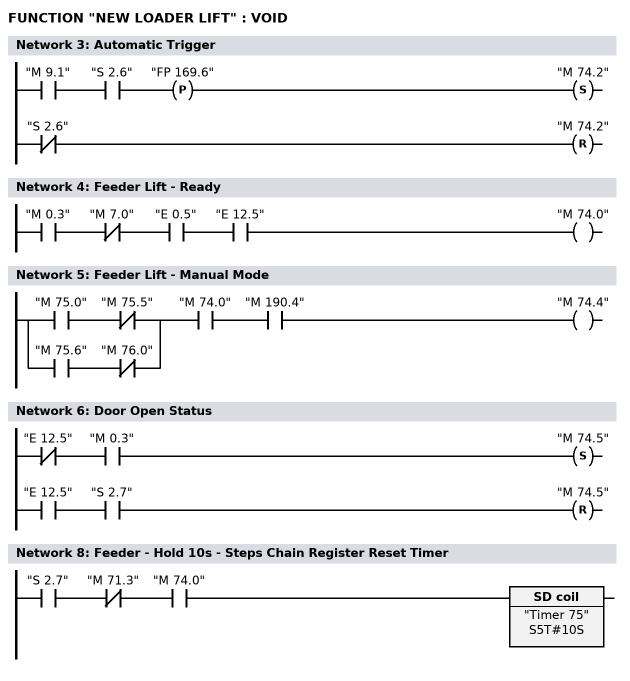

      O     "M 9.1";
      A     "S 2.6";
      FP    "FP 169.6";
      S     "M 74.2";
//;
      AN    "S 2.6";
      R     "M 74.2";
NETWORK
TITLE =Feeder Lift - Ready

      A     "M 0.3";
      AN    "M 7.0";
      A     "E 0.5";
      A     "E 12.5";
      =     "M 74.0";
NETWORK
TITLE =Feeder Lift - Manual Mode

      A(    ;
      A     "M 75.0";
      AN    "M 75.5";
      O     ;
      A     "M 75.6";
      AN    "M 76.0";
      )     ;
      A     "M 74.0";
      A     "M 190.4";
      =     "M 74.4";
NETWORK
TITLE =Door Open Status

      AN    "E 12.5";
      A     "M 0.3";
      S     "M 74.5";
//;
      A     "E 12.5";
      A     "S 2.7";
      R     "M 74.5";
NETWORK
TITLE =Fault Reset Status        X121     transfered to FC 212 Net 79
//      A(
//      O     "M 54.7"
//      O     "M 66.7"
//      O     "M 86.7"
//      )
//      A     "M 145.0"
//      O     "M 74.5"
//      O     "Timer 0"
//      =     "H 40.3"
//
//is transfered to FC 212 Net 79


NETWORK
TITLE =Feeder - Hold 10s - Steps Chain Register Reset Timer

      A     "S 2.7";
      AN    "M 71.3";
      A     "M 74.0";
      L     S5T#10S;
      SD    "Timer 75";
NETWORK
TITLE =Feeder - All Register Reset

      A(    ;
      A     "M 190.4";
      A     "M 171.4";
      A     "M 171.5";
      O     "Timer 75";
      )     ;
      A     "M 74.0";
      JC    M001;
      JU    M002;

M001: L     2#0;
      T     "MW 71";
      T     "MW 75";

M002: NOP   0;
NETWORK
TITLE =Step 16N1 - Power On
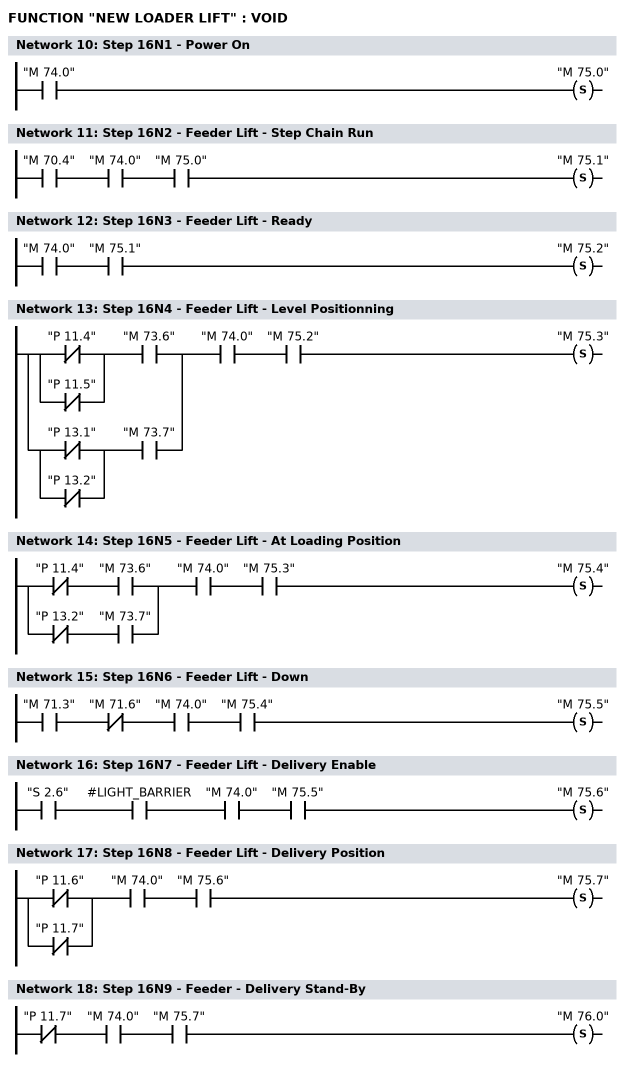

      A     "M 74.0";
      S     "M 75.0";
NETWORK
TITLE =Step 16N2 - Feeder Lift - Step Chain Run

      A     "M 70.4";
      A     "M 74.0";
      A     "M 75.0";
      S     "M 75.1";
NETWORK
TITLE =Step 16N3 - Feeder Lift - Ready

      A     "M 74.0";
      A     "M 75.1";
      S     "M 75.2";
NETWORK
TITLE =Step 16N4 - Feeder Lift - Level Positionning

      A(    ;
      A(    ;
      ON    "P 11.4";
      ON    "P 11.5";
      )     ;
      A     "M 73.6";
      O     ;
      A(    ;
      ON    "P 13.1";
      ON    "P 13.2";
      )     ;
      A     "M 73.7";
      )     ;
      A     "M 74.0";
      A     "M 75.2";
      S     "M 75.3";
NETWORK
TITLE =Step 16N5 - Feeder Lift - At Loading Position

      A(    ;
      AN    "P 11.4";
      A     "M 73.6";
      O     ;
      AN    "P 13.2";
      A     "M 73.7";
      )     ;
      A     "M 74.0";
      A     "M 75.3";
      S     "M 75.4";
NETWORK
TITLE =Step 16N6 - Feeder Lift - Down

      A     "M 71.3";
      AN    "M 71.6";
      A     "M 74.0";
      A     "M 75.4";
      S     "M 75.5";
NETWORK
TITLE =Step 16N7 - Feeder Lift - Delivery Enable

      A     "S 2.6";
      A     #LIGHT_BARRIER;
      A     "M 74.0";
      A     "M 75.5";
      S     "M 75.6";
NETWORK
TITLE =Step 16N8 - Feeder Lift - Delivery Position

      A(    ;
      ON    "P 11.6";
      ON    "P 11.7";
      )     ;
      A     "M 74.0";
      A     "M 75.6";
      S     "M 75.7";
NETWORK
TITLE =Step 16N9 - Feeder - Delivery Stand-By

      AN    "P 11.7";
      A     "M 74.0";
      A     "M 75.7";
      S     "M 76.0";
NETWORK
TITLE =Feeder Lift Steps Chain Reset by Feeder Fingers (MW71)

      A     "M 76.0";
      AN    "M 76.1";
      A(    ;
      ON    "M 71.2";
      O     "M 72.2";
      )     ;
      A     "M 74.0";
      JC    M003;
      JU    M004;

M003: L     2#0;
      T     "MW 75";

M004: NOP   0;
NETWORK
TITLE =Step 16N10 - Feeder Hold Operation (Stop) 1
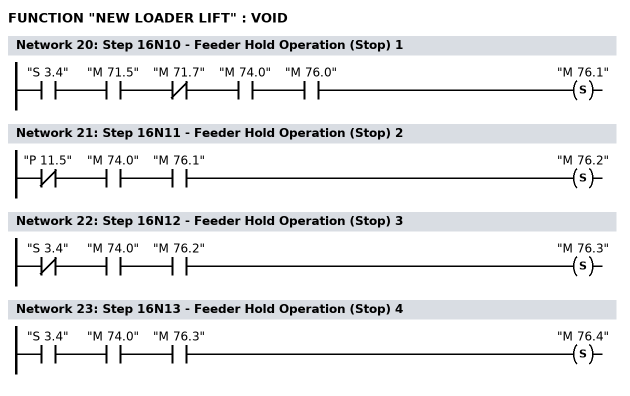

      A     "S 3.4";
      A     "M 71.5";
      AN    "M 71.7";
      A     "M 74.0";
      A     "M 76.0";
      S     "M 76.1";
NETWORK
TITLE =Step 16N11 - Feeder Hold Operation (Stop) 2

      AN    "P 11.5";
      A     "M 74.0";
      A     "M 76.1";
      S     "M 76.2";
NETWORK
TITLE =Step 16N12 - Feeder Hold Operation (Stop) 3

      AN    "S 3.4";
      A     "M 74.0";
      A     "M 76.2";
      S     "M 76.3";
NETWORK
TITLE =Step 16N13 - Feeder Hold Operation (Stop) 4

      A     "S 3.4";
      A     "M 74.0";
      A     "M 76.3";
      S     "M 76.4";
NETWORK
TITLE =Step 16N14 - Feeder Hold Operation (Stop) 4 - Fill MB76

      A     "M 76.4";
      A     "M 74.0";
      JC    M005;
      JU    M006;

M005: L     2#11111100000000;
      T     "MW 75";

M006: NOP   0;
NETWORK
TITLE =Packets Movements - UpDate
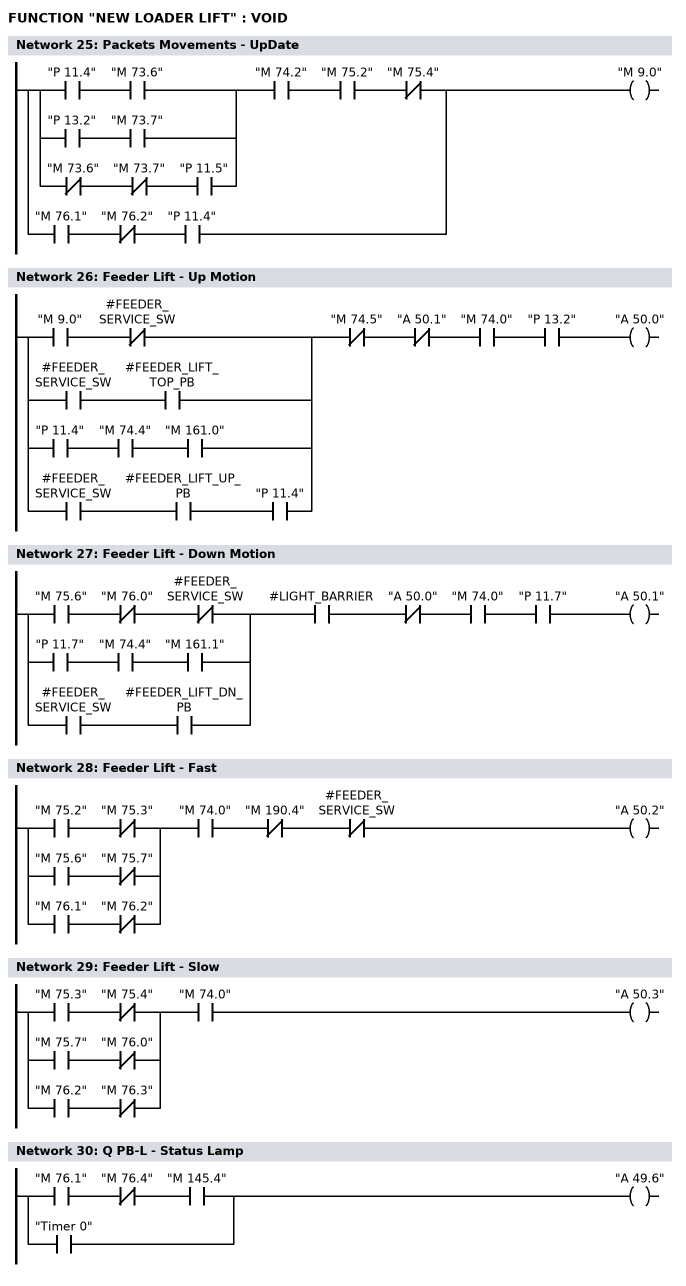

      A(    ;
      A     "P 11.4";
      A     "M 73.6";
      O     ;
      A     "P 13.2";
      A     "M 73.7";
      O     ;
      AN    "M 73.6";
      AN    "M 73.7";
      A     "P 11.5";
      )     ;
      A     "M 74.2";
      A     "M 75.2";
      AN    "M 75.4";
      O     ;
      A     "M 76.1";
      AN    "M 76.2";
      A     "P 11.4";
      =     "M 9.0";
NETWORK
TITLE =Feeder Lift - Up Motion

      A(    ;
      A     "M 9.0";
      AN    #FEEDER_SERVICE_SW;
      O     ;
      A     #FEEDER_SERVICE_SW;
      A     #FEEDER_LIFT_TOP_PB;

      O     ;
      A     "P 11.4";
      A     "M 74.4";
      A     "M 161.0";

      O     ;
      A     #FEEDER_SERVICE_SW;
      A     #FEEDER_LIFT_UP_PB;
      A     "P 11.4";
      )     ;
      AN    "M 74.5";
      AN    "A 50.1";
      A     "M 74.0";
      A     "P 13.2";
      =     "A 50.0";
NETWORK
TITLE =Feeder Lift - Down Motion

      A(    ;
      A     "M 75.6";
      AN    "M 76.0";
      AN    #FEEDER_SERVICE_SW;

      O     ;
      A     "P 11.7";
      A     "M 74.4";
      A     "M 161.1";

      O     ;
      A     #FEEDER_SERVICE_SW;
      A     #FEEDER_LIFT_DN_PB;
      )     ;
      A     #LIGHT_BARRIER;
      AN    "A 50.0";
      A     "M 74.0";
      A     "P 11.7";
      =     "A 50.1";
NETWORK
TITLE =Feeder Lift - Fast

      A(    ;
      A     "M 75.2";
      AN    "M 75.3";
      O     ;
      A     "M 75.6";
      AN    "M 75.7";
      O     ;
      A     "M 76.1";
      AN    "M 76.2";
      )     ;
      A     "M 74.0";
      AN    "M 190.4";
      AN    #FEEDER_SERVICE_SW;
      =     "A 50.2";
NETWORK
TITLE =Feeder Lift - Slow

      A(    ;
      A     "M 75.3";
      AN    "M 75.4";
      O     ;
      A     "M 75.7";
      AN    "M 76.0";
      O     ;
      A     "M 76.2";
      AN    "M 76.3";
      )     ;
      A     "M 74.0";
      =     "A 50.3";
NETWORK
TITLE =Q PB-L - Status Lamp

      A     "M 76.1";
      AN    "M 76.4";
      A     "M 145.4";
      O     "Timer 0";
      =     "A 49.6";
END_FUNCTION

FUNCTION "NEW C21 - LINK 1 HI" : VOID
TITLE =NEW FC978 (was FC1078) - Conveyor 21 - Link 1H Pos. 13 High Leve
//
//v0.1 2026-11-19: clearing trigger M9.3 only if pivot HIGH (P15.0).
NAME : POS_13_H
VERSION : 0.1


VAR_TEMP
  MAIN_SERVICE_2_SW : BOOL ;
  SERVICE_RUN : BOOL ;
  INITIALISATION : BOOL ;
  BARRIER_BLINKER : BOOL ;
END_VAR
BEGIN
NETWORK
TITLE =Conveyor 21 - Service

      A     "HMI_DB".ALL_SERVICE_ENABLE_SW;
      A     "HMI_DB".CONVEYOR_21_SERVICE_SW;
      A     "HMI_DB".SERVICE_SW_2_STATUS;
      =     #MAIN_SERVICE_2_SW;
//;
      A     #MAIN_SERVICE_2_SW;
      O     "M 78.7";
      JNB   CO21;
//;
      A     "HMI_DB".HMI_CONVEYOR_21_TEST_SSW;
      AN    "A 48.0";
      =     #SERVICE_RUN;
      S     "DB UTILITY".Conveyor_10_Disable;
      S     "DB UTILITY".Pivot_Disable;
//;
      A     "HMI_DB".SERVICE_INIT_PB;
      =     #INITIALISATION;
//;
      AN    #MAIN_SERVICE_2_SW;
      R     "HMI_DB".HMI_CONVEYOR_21_TEST_SSW;
      R     "DB UTILITY".Conveyor_10_Disable;
      R     "DB UTILITY".Pivot_Disable;

CO21: R     #SERVICE_RUN;
      R     #INITIALISATION; // Fix: temp not written when service is off
      FP    "FP 148.3";
      =     "M 78.7";
NETWORK
TITLE =Power Enable
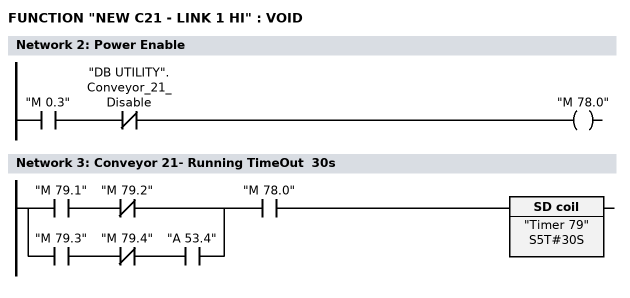

      A     "M 0.3";
      AN    "DB UTILITY".Conveyor_21_Disable;
      =     "M 78.0";
NETWORK
TITLE =Conveyor 21- Running TimeOut  30s

      A(    ;
      A     "M 79.1";
      AN    "M 79.2";
      O     ;
      A     "M 79.3";
      AN    "M 79.4";
      A     "A 53.4";
      )     ;
      A     "M 78.0";
      L     S5T#30S;
      SD    "Timer 79"; // C21 TimeOut
NETWORK
TITLE =Steps Register - Reset

      A(    ;
      A     "M 79.1"; // Filling Step
      AN    "M 79.2"; // Filling Step - Done
      A     "Timer 79"; // C21 TimeOut
      O     "M 79.4";
      O     #INITIALISATION;
      O     "DB UTILITY".Conveyor_21_Disable;
      )     ;
      A     "M 78.0";
      JC    M001;
      JU    M002;

M001: L     W#16#0;
      T     "MW 79"; // Step Register - Reset
      T     "MB 81"; // Step Register - Reset

M002: NOP   0;
NETWORK
TITLE =Step 22N1 - Power ON
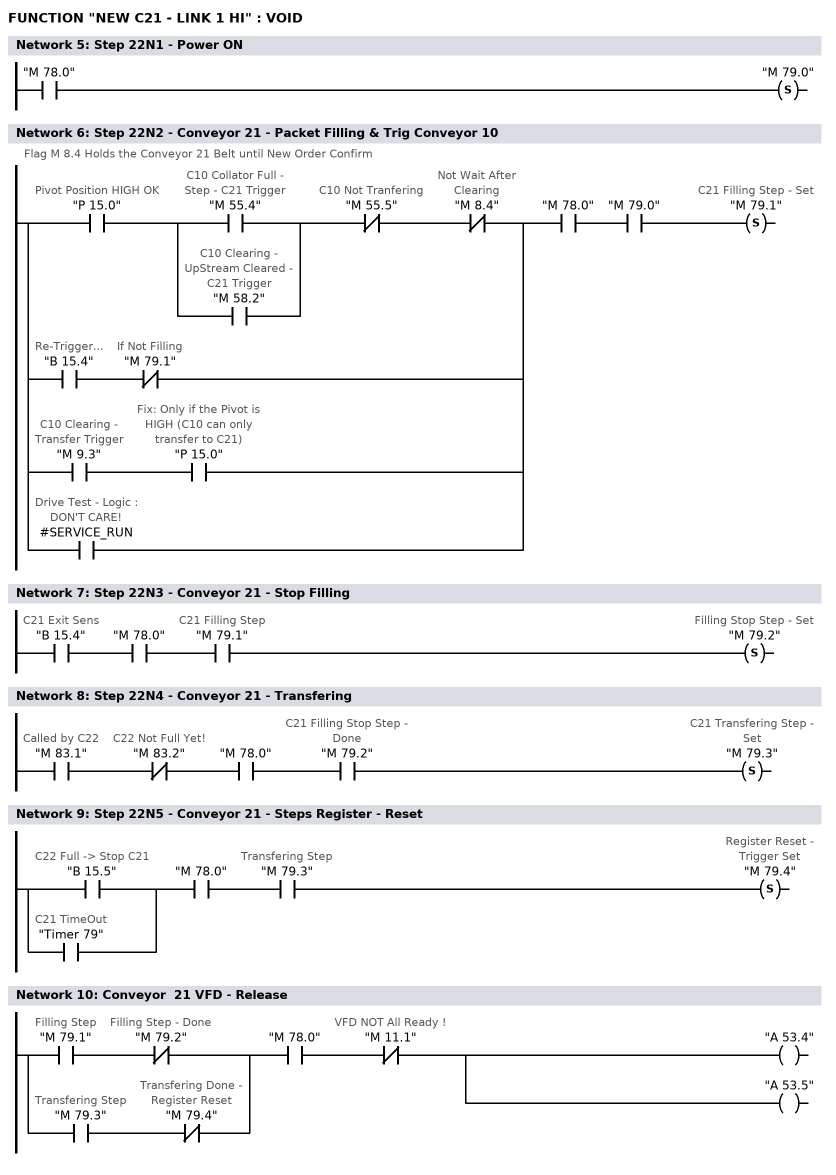

      A     "M 78.0";
      S     "M 79.0";
NETWORK
TITLE =Step 22N2 - Conveyor 21 - Packet Filling & Trig Conveyor 10
//Flag M 8.4 Holds the Conveyor 21 Belt until New Order Confirm
      A(    ;
      A     "P 15.0"; // Pivot Position HIGH OK
      A(    ;
      O     "M 55.4"; // C10 Collator Full - Step - C21 Trigger
      O     "M 58.2"; // C10 Clearing - UpStream Cleared - C21 Trigger
      )     ;
      AN    "M 55.5"; // C10 Not Tranfering
      AN    "M 8.4"; // Not Wait After Clearing
      O     ;
      A     "B 15.4"; // Re-Trigger...
      AN    "M 79.1"; // If Not Filling
      O     ;
      A     "M 9.3"; // C10 Clearing - Transfer Trigger
      A     "P 15.0"; // Fix: Only if the Pivot is HIGH (C10 can only transfer to C21)
      )     ;
      O     #SERVICE_RUN; // Drive Test - Logic : DON'T CARE!
      A     "M 78.0";
      A     "M 79.0";
      S     "M 79.1"; // C21 Filling Step - Set
NETWORK
TITLE =Step 22N3 - Conveyor 21 - Stop Filling

      A     "B 15.4"; // C21 Exit Sens
      A     "M 78.0";
      A     "M 79.1"; // C21 Filling Step
      S     "M 79.2"; // Filling Stop Step - Set
NETWORK
TITLE =Step 22N4 - Conveyor 21 - Transfering

      A     "M 83.1"; // Called by C22
      AN    "M 83.2"; // C22 Not Full Yet!
      A     "M 78.0";
      A     "M 79.2"; // C21 Filling Stop Step - Done
      S     "M 79.3"; // C21 Transfering Step - Set
NETWORK
TITLE =Step 22N5 - Conveyor 21 - Steps Register - Reset

      A(    ;
      O     "B 15.5"; // C22 Full -> Stop C21
      O     "Timer 79"; // C21 TimeOut
      )     ;
      A     "M 78.0";
      A     "M 79.3"; // Transfering Step
      S     "M 79.4"; // Register Reset - Trigger Set
NETWORK
TITLE =Conveyor  21 VFD - Release

      A(    ;
      A     "M 79.1"; // Filling Step
      AN    "M 79.2"; // Filling Step - Done
      O     ;
      A     "M 79.3"; // Transfering Step
      AN    "M 79.4"; // Transfering Done - Register Reset
      )     ;
      A     "M 78.0";
      AN    "M 11.1"; // VFD NOT All Ready !
      =     "A 53.4";
      =     "A 53.5";
END_FUNCTION

FUNCTION "NEW C22 - LINK 2 HI" : VOID
TITLE =NEW FC982 (was FC1082) - Conveyor 22 - Link 2H Pos. 14 High Leve
//
NAME : POS_14_H
VERSION : 0.0


VAR_TEMP
  MAIN_SERVICE_2_SW : BOOL ;
  SERVICE_RUN : BOOL ;
END_VAR
BEGIN
NETWORK
TITLE =Conveyor 22 - Service

      A     "HMI_DB".ALL_SERVICE_ENABLE_SW;
      A     "HMI_DB".CONVEYOR_21_SERVICE_SW;
      A     "HMI_DB".SERVICE_SW_2_STATUS;
      =     #MAIN_SERVICE_2_SW;
//;
      A     #MAIN_SERVICE_2_SW;
      O     "M 82.7";
      JNB   CO22;
//;
      A     "HMI_DB".HMI_CONVEYOR_22_TEST_SSW;
      =     #SERVICE_RUN;
//;
      AN    #MAIN_SERVICE_2_SW;
      R     "HMI_DB".HMI_CONVEYOR_22_TEST_SSW;

CO22: R     #SERVICE_RUN;
      FP    "FP 148.4";
      =     "M 82.7";
NETWORK
TITLE =Power Enable
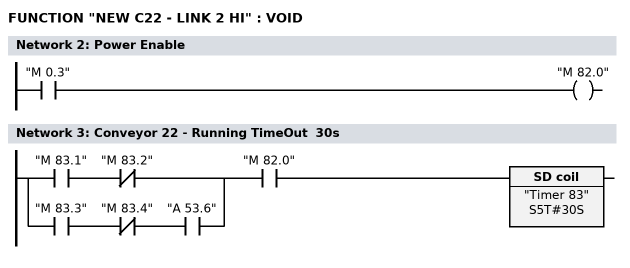

      A     "M 0.3";
      =     "M 82.0";
NETWORK
TITLE =Conveyor 22 - Running TimeOut  30s

      A(    ;
      A     "M 83.1";
      AN    "M 83.2";
      O     ;
      A     "M 83.3";
      AN    "M 83.4";
      A     "A 53.6";
      )     ;
      A     "M 82.0";
      L     S5T#30S;
      SD    "Timer 83";
NETWORK
TITLE =Conveyor 22 - Steps Register - Reset

      A(    ;
      A     "M 83.1";
      AN    "M 83.2";
      A     "Timer 83";
      O     "M 83.4";
      )     ;
      A     "M 82.0";
      JC    M001;
      JU    M002;

M001: L     W#16#0;
      T     "MW 83";
      T     "MB 85";

M002: NOP   0;
NETWORK
TITLE =Step 23N1 - Power On
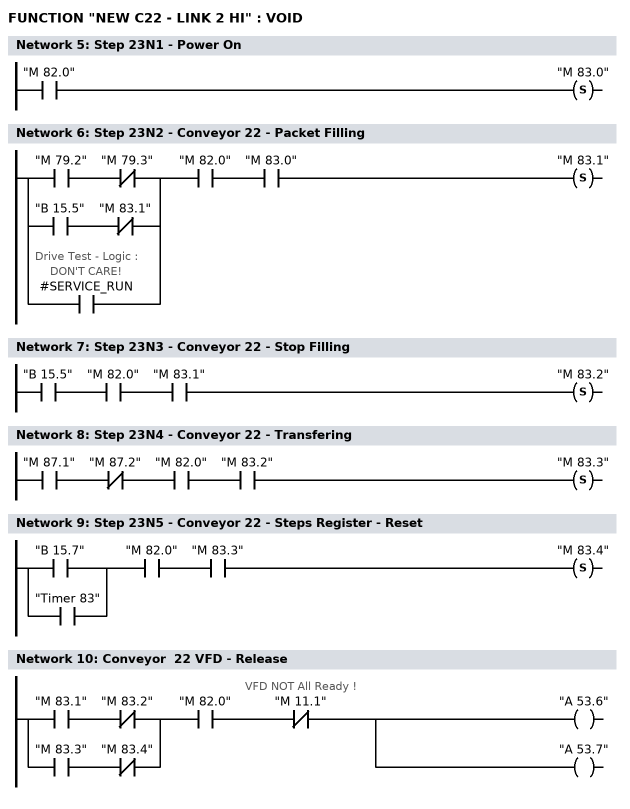

      A     "M 82.0";
      S     "M 83.0";
NETWORK
TITLE =Step 23N2 - Conveyor 22 - Packet Filling

      A(    ;
      A     "M 79.2";
      AN    "M 79.3";
      O     ;
      A     "B 15.5";
      AN    "M 83.1";
      )     ;
      O     #SERVICE_RUN; // Drive Test - Logic : DON'T CARE!
      A     "M 82.0";
      A     "M 83.0";
      S     "M 83.1";
NETWORK
TITLE =Step 23N3 - Conveyor 22 - Stop Filling

      A     "B 15.5";
      A     "M 82.0";
      A     "M 83.1";
      S     "M 83.2";
NETWORK
TITLE =Step 23N4 - Conveyor 22 - Transfering

      A     "M 87.1";
      AN    "M 87.2";
      A     "M 82.0";
      A     "M 83.2";
      S     "M 83.3";
NETWORK
TITLE =Step 23N5 - Conveyor 22 - Steps Register - Reset

      A(    ;
      O     "B 15.7";
      O     "Timer 83";
      )     ;
      A     "M 82.0";
      A     "M 83.3";
      S     "M 83.4";
NETWORK
TITLE =Conveyor  22 VFD - Release

      A(    ;
      A     "M 83.1";
      AN    "M 83.2";
      O     ;
      A     "M 83.3";
      AN    "M 83.4";
      )     ;
      A     "M 82.0";
      AN    "M 11.1"; // VFD NOT All Ready !
      =     "A 53.6";
      =     "A 53.7";
END_FUNCTION

FUNCTION "NEW C23 - DELIV. HI" : VOID
TITLE =NEW FC986 (was FC1086) - Conveyor 23 - Delivery Second Level
//
NAME : POS_15_H
VERSION : 0.0


VAR_TEMP
  MAIN_SERVICE_2_SW : BOOL ;
  SERVICE_RUN : BOOL ;
END_VAR
BEGIN
NETWORK
TITLE =Conveyor 23 - Service

      A     "HMI_DB".ALL_SERVICE_ENABLE_SW;
      A     "HMI_DB".CONVEYOR_21_SERVICE_SW;
      A     "HMI_DB".SERVICE_SW_2_STATUS;
      =     #MAIN_SERVICE_2_SW;
//;
      A     #MAIN_SERVICE_2_SW;
      O     "M 86.1";
      JNB   CO23;
//;
      A     "HMI_DB".HMI_CONVEYOR_23_TEST_SSW;
      =     #SERVICE_RUN;
//;
      AN    #MAIN_SERVICE_2_SW;
      R     "HMI_DB".HMI_CONVEYOR_23_TEST_SSW;

CO23: R     #SERVICE_RUN;
      FP    "FP 149.3";
      =     "M 86.1";
NETWORK
TITLE =Delivery Conveyor 23 - Running TimeOut  30s
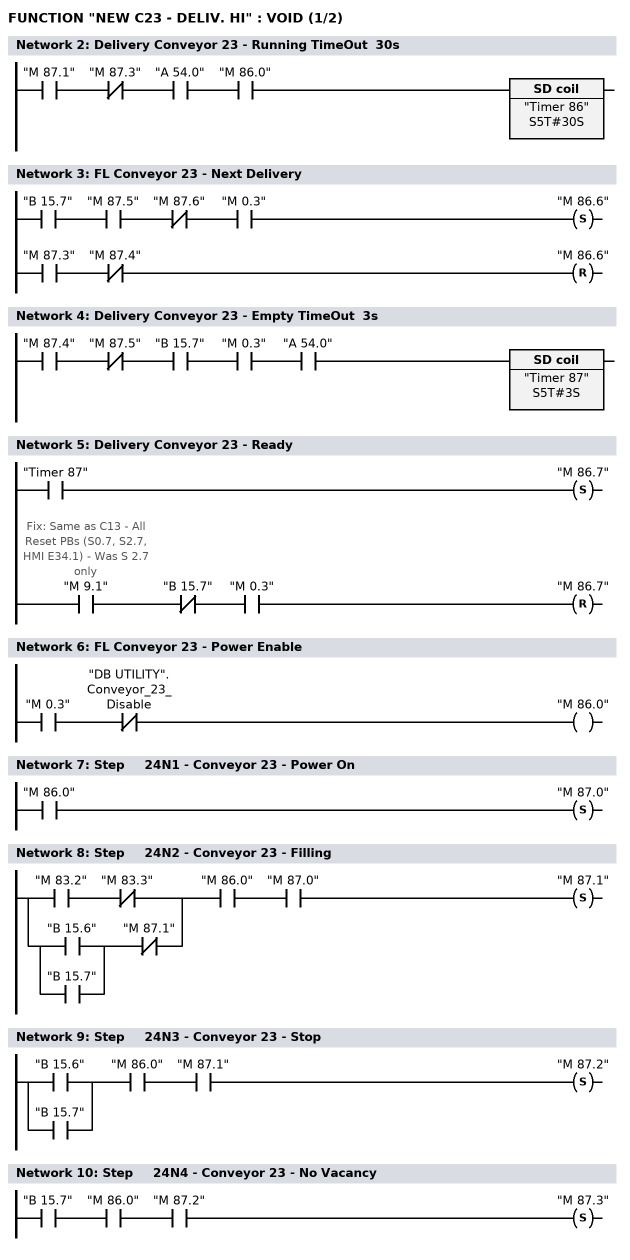

      A     "M 87.1";
      AN    "M 87.3";
      A     "A 54.0";
      A     "M 86.0";
      L     S5T#30S;
      SD    "Timer 86";
NETWORK
TITLE =FL Conveyor 23 - Next Delivery

      A     "B 15.7";
      A     "M 87.5";
      AN    "M 87.6";
      A     "M 0.3";
      S     "M 86.6";
//;
      A     "M 87.3";
      AN    "M 87.4";
      R     "M 86.6";
NETWORK
TITLE =Delivery Conveyor 23 - Empty TimeOut  3s

      A     "M 87.4";
      AN    "M 87.5";
      A     "B 15.7";
      A     "M 0.3";
      A     "A 54.0";
      L     S5T#3S;
      SD    "Timer 87";
NETWORK
TITLE =Delivery Conveyor 23 - Ready

      A     "Timer 87";
      S     "M 86.7";
//;
      A     "M 9.1"; // Fix: Same as C13 - All Reset PBs (S0.7, S2.7, HMI E34.1) - Was S 2.7 only
      AN    "B 15.7";
      A     "M 0.3";
      R     "M 86.7";
NETWORK
TITLE =FL Conveyor 23 - Power Enable

      A     "M 0.3";
      AN    "DB UTILITY".Conveyor_23_Disable;
      =     "M 86.0";
NETWORK
TITLE =Step     24N1 - Conveyor 23 - Power On

      A     "M 86.0";
      S     "M 87.0";
NETWORK
TITLE =Step     24N2 - Conveyor 23 - Filling

      A(    ;
      A     "M 83.2";
      AN    "M 83.3";
      O     ;
      A(    ;
      O     "B 15.6";
      O     "B 15.7";
      )     ;
//      O     #SERVICE_RUN
      AN    "M 87.1";
      )     ;
      A     "M 86.0";
      A     "M 87.0";
      S     "M 87.1";
NETWORK
TITLE =Step     24N3 - Conveyor 23 - Stop

      A(    ;
      O     "B 15.6";
      O     "B 15.7";
      )     ;
      A     "M 86.0";
      A     "M 87.1";
      S     "M 87.2";
NETWORK
TITLE =Step     24N4 - Conveyor 23 - No Vacancy

      A     "B 15.7";
      A     "M 86.0";
      A     "M 87.2";
      S     "M 87.3";
NETWORK
TITLE =Step     24N5 - Conveyor 23 - Delivery
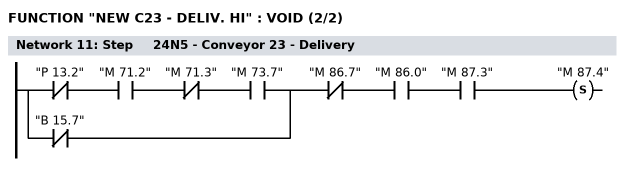

      A(    ;
      AN    "P 13.2";
      A     "M 71.2";
      AN    "M 71.3";
      A     "M 73.7";
      ON    "B 15.7";
      )     ;
      AN    "M 86.7";
      A     "M 86.0";
      A     "M 87.3";
      S     "M 87.4";
NETWORK
TITLE =Write 1 to Steps 0-3 Byte Register MB87

      A(    ;
      O     "M 86.6";
      O     "M 86.7";
      )     ;
      A     "M 87.4";
      A     "M 86.0";
      JC    M001;
      JU    M002;

M001: L     2#1111;
      T     "MB 87";

M002: NOP   0;
NETWORK
TITLE =Step     24N6 - Conveyor 23 - Delivery Done
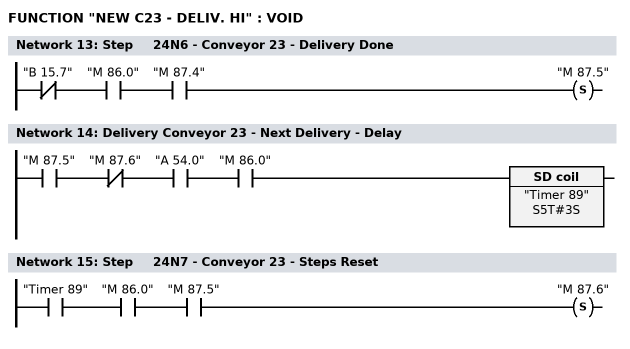

      AN    "B 15.7";
      A     "M 86.0";
      A     "M 87.4";
      S     "M 87.5";
NETWORK
TITLE =Delivery Conveyor 23 - Next Delivery - Delay

      A     "M 87.5";
      AN    "M 87.6";
      A     "A 54.0";
      A     "M 86.0";
      L     S5T#3S;
      SD    "Timer 89";
NETWORK
TITLE =Step     24N7 - Conveyor 23 - Steps Reset

      A     "Timer 89";
      A     "M 86.0";
      A     "M 87.5";
      S     "M 87.6";
NETWORK
TITLE =Steps Register - Reset

      A(    ;
      O     "M 87.6";
      O     "Timer 86";
      )     ;
      A     "M 86.0";
      JC    M003;
      JU    M004;

M003: L     2#0;
      T     "MW 87";

M004: NOP   0;
NETWORK
TITLE =Conveyor  23 VFD - Release
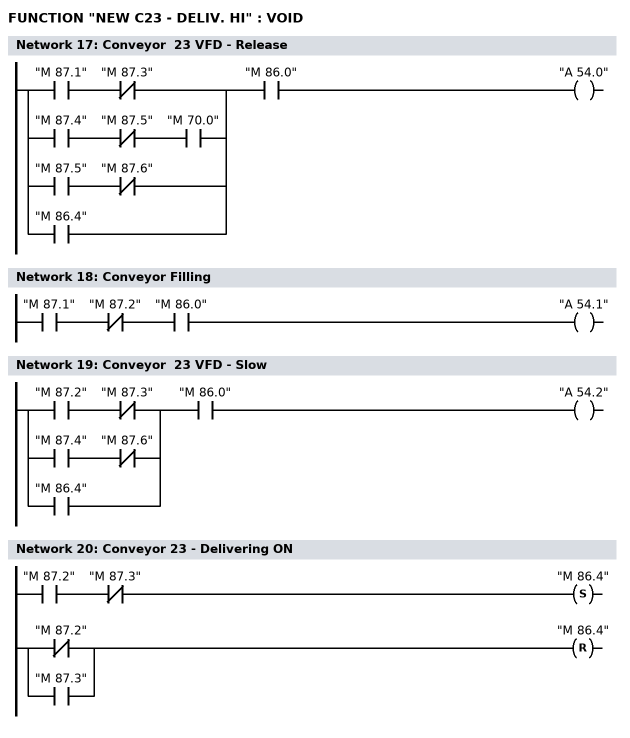

      A(    ;
      A     "M 87.1";
      AN    "M 87.3";
      O     ;
      A     "M 87.4";
      AN    "M 87.5";
      A     "M 70.0";
      O     ;
      A     "M 87.5";
      AN    "M 87.6";
      O     "M 86.4";
      )     ;
      A     "M 86.0";
      =     "A 54.0";
NETWORK
TITLE =Conveyor Filling

      A     "M 87.1";
      AN    "M 87.2";
      A     "M 86.0";
      =     "A 54.1";
NETWORK
TITLE =Conveyor  23 VFD - Slow

      A(    ;
      A     "M 87.2";
      AN    "M 87.3";
      O     ;
      A     "M 87.4";
      AN    "M 87.6";
      O     "M 86.4";
      )     ;
      A     "M 86.0";
      =     "A 54.2";
NETWORK
TITLE =Conveyor 23 - Delivering ON

      A     "M 87.2";
      AN    "M 87.3";
      S     "M 86.4";
      A(    ;
      ON    "M 87.2";
      O     "M 87.3";
      )     ;
      R     "M 86.4";
END_FUNCTION

FUNCTION "LIGHT BAR" : VOID
TITLE =Light Bar
VERSION : 0.1


VAR_TEMP
  BARRIER_BLINKER : BOOL ;	//Feeder Safety Light Barrier
  STATUS_BLANKER : BOOL ;
  CLEARING_BLINKER : BOOL ;
END_VAR
BEGIN
NETWORK
TITLE =Light Barrier - Blinker
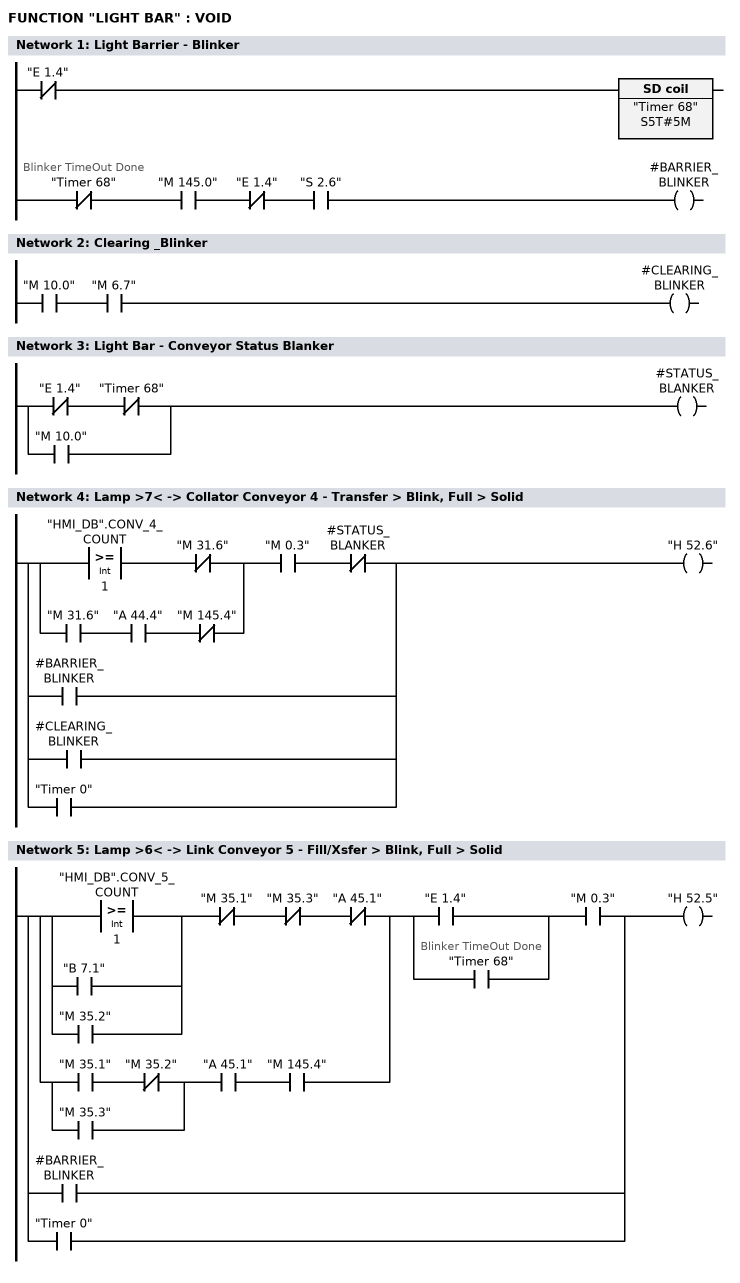

      ON    "E 1.4";
      L     S5T#5M;
      SD    "Timer 68"; // Blinker TimeOut Start
//;
      A(    ;
      AN    "Timer 68"; // Blinker TimeOut Done
      A     "M 145.0";
      )     ;
      AN    "E 1.4";
      A     "S 2.6";
      =     #BARRIER_BLINKER;
NETWORK
TITLE =Clearing _Blinker

      A     "M 10.0";
      A     "M 6.7";
      =     #CLEARING_BLINKER;
NETWORK
TITLE =Light Bar - Conveyor Status Blanker

      AN    "E 1.4";
      AN    "Timer 68";
      O     "M 10.0";
      =     #STATUS_BLANKER;
NETWORK
TITLE =Lamp >7< -> Collator Conveyor 4 - Transfer > Blink, Full > Solid

      A(    ;

      A(    ; // Solid
      A(    ;
      L     "HMI_DB".CONV_4_COUNT;
      L     1;
      >=I   ;
      )     ;
      AN    "M 31.6";
      )     ; // Solid

      O     ;

      A(    ; // Blink
      A     "M 31.6";
      A     "A 44.4";
      AN    "M 145.4";
      )     ; // Blink

      )     ;
      A     "M 0.3";
      AN    #STATUS_BLANKER;
      O     #BARRIER_BLINKER;
      O     #CLEARING_BLINKER;
      O     "Timer 0";
      =     "H 52.6";
NETWORK
TITLE =Lamp >6< -> Link Conveyor 5 - Fill/Xsfer > Blink, Full > Solid

      A(    ;

      A(    ; // Solid
      A(    ;
      A(    ;
      L     "HMI_DB".CONV_5_COUNT;
      L     1;
      >=I   ;
      )     ;
      O     "B 7.1";
      )     ;
      O     "M 35.2";
      AN    "M 35.1";
      AN    "M 35.3";
      AN    "A 45.1";
      )     ; // Solid

      O     ;

      A(    ; // Blink
      A(    ;
      A     "M 35.1";
      AN    "M 35.2";
      O     ;
      A     "M 35.3";
      )     ;
      A     "A 45.1";
      A     "M 145.4";
      )     ; // Blink

      )     ;
      A(    ;
      A     "E 1.4";
      O     "Timer 68"; // Blinker TimeOut Done
      )     ;
      A     "M 0.3";
      O     #BARRIER_BLINKER;
      O     "Timer 0";
      =     "H 52.5";
NETWORK
TITLE =Lamp >5< -> Delivery Conveyor 6 - Fill > Blink, Full > Solid

      A(    ;

      A(    ; // Solid
      A(    ;
      A(    ;
      L     "HMI_DB".CONV_6_COUNT;
      L     1;
      >=I   ;
      )     ;
      O     "B 7.2";
      )     ;
      O     "M 39.2";
      AN(   ;
      A     "M 39.1";
      AN    "M 39.2";
      )     ;
      AN    "A 45.4";
      )     ; // Solid

      O     ;

      A(    ; // Blink
      A     "M 39.1";
      AN    "M 39.2";
      A     "A 45.4";
      AN    "M 145.4";
      )     ; // Blink

      )     ;
      A(    ;
      A     "E 1.4";
      O     "Timer 68"; // Blinker TimeOut Done
      )     ;
      A     "M 0.3";
      O     #BARRIER_BLINKER;
      O     "Timer 0";
      =     "H 52.4";
NETWORK
TITLE =Lamp >4< -> Pivot 10 -> 11L/21H - Fill > Blink, Full > Solid
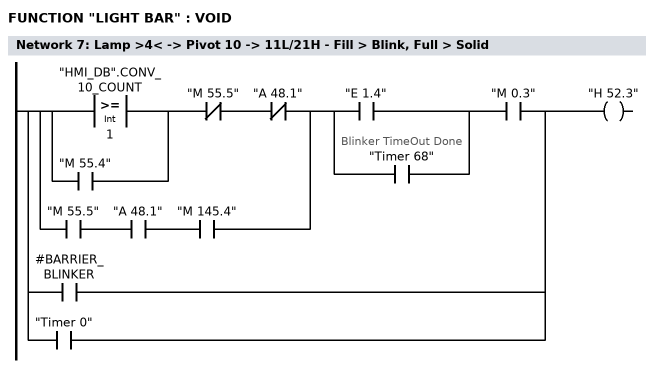

      A(    ;

      A(    ; // Solid
      A(    ;
      L     "HMI_DB".CONV_10_COUNT;
      L     1;
      >=I   ;
      )     ;
      O     "M 55.4";
      AN    "M 55.5";
      AN    "A 48.1";
      )     ; // Solid

      O     ;

      A(    ; // Blink
      A     "M 55.5";
      A     "A 48.1";
      A     "M 145.4";
      )     ; // Blink

      )     ;
      A(    ;
      A     "E 1.4";
      O     "Timer 68"; // Blinker TimeOut Done
      )     ;
      A     "M 0.3";
      O     #BARRIER_BLINKER;
      O     "Timer 0";
      =     "H 52.3";
NETWORK
TITLE =Lamp >3< -> Link Conveyors 11L/21H - Fill > Blink, Full > Solid

      A(    ;

      A(    ; // Solid
      A(    ;
      A(    ;
      A(    ;
      L     "HMI_DB".CONV_11_COUNT;
      L     "HMI_DB".CONV_21_COUNT;
      +I    ;
      L     1;
      >=I   ;
      )     ;
      O     "B 10.7";
      O     "B 15.4";
      )     ;
      O     "M 59.2";
      O     "M 79.2";
      )     ;
      AN(   ;
      A     "M 59.1";
      AN    "M 59.2";
      )     ;
      AN(   ;
      A     "M 79.1";
      AN    "M 79.2";
      )     ;
      AN    "M 59.3";
      AN    "M 79.3";
      AN    "A 48.3";
      AN    "A 53.4";
      )     ; // Solid

      O     ;

      A(    ; // Blink
      A(    ;
      A(    ;
      A     "M 59.1";
      AN    "M 59.2";
      O     ;
      A     "M 79.1";
      AN    "M 79.2";
      )     ;
      O     ;
      A(    ;
      A     "M 59.3";
      O     "M 79.3";
      )     ;
      )     ;
      A(    ;
      O     "A 48.3";
      O     "A 53.4";
      )     ;
      AN    "M 145.4";
      )     ; // Blink

      )     ;
      A(    ;
      A     "E 1.4";
      O     "Timer 68"; // Blinker TimeOut Done
      )     ;
      A     "M 0.3";
      O     #BARRIER_BLINKER;
      O     "Timer 0";
      =     "H 52.2";

NETWORK
TITLE =Lamp >2< -> Link Conveyors 12L/22H - Fill > Blink, Full > Solid

      A(    ;

      A(    ; // Solid
      A(    ;
      A(    ;
      A(    ;
      L     "HMI_DB".CONV_12_COUNT;
      L     "HMI_DB".CONV_22_COUNT;
      +I    ;
      L     1;
      >=I   ;
      )     ;
      O     "B 11.0";
      O     "B 15.5";
      )     ;
      O     "M 63.2";
      O     "M 83.2";
      )     ;
      AN(   ;
      A     "M 63.1";
      AN    "M 63.2";
      )     ;
      AN(   ;
      A     "M 83.1";
      AN    "M 83.2";
      )     ;
      AN    "M 63.3";
      AN    "M 83.3";
      AN    "A 48.6";
      AN    "A 53.6";
      )     ; // Solid

      O     ;

      A(    ; // Blink
      A(    ;
      A(    ;
      A     "M 63.1";
      AN    "M 63.2";
      O     ;
      A     "M 83.1";
      AN    "M 83.2";
      )     ;
      O     ;
      A(    ;
      A     "M 63.3";
      O     "M 83.3";
      )     ;
      )     ;
      A(    ;
      O     "A 48.6";
      O     "A 53.6";
      )     ;
      A     "M 145.4";
      )     ; // Blink

      )     ;
      A(    ;
      A     "E 1.4";
      O     "Timer 68"; // Blinker TimeOut Done
      )     ;
      A     "M 0.3";
      O     #BARRIER_BLINKER;
      O     "Timer 0";
      =     "H 52.1";

NETWORK
TITLE =Lamp >1< -> Output Conveyors 13L/23H - Fill > Blink,Full > Solid

      A(    ; // Solid

      A(    ;
      L     "HMI_DB".CONV_13_COUNT;
      L     "HMI_DB".CONV_23_COUNT;
      +I    ;
      L     1;
      >=I   ;
      )     ;
      O     "B 11.2";
      O     "B 15.7";
      )     ; // Solid

      A(    ;
      A     "E 1.4";
      O     "Timer 68"; // Blinker TimeOut Done
      )     ;
      A     "M 0.3";
      AN    #STATUS_BLANKER;
      O     #BARRIER_BLINKER;
      O     #CLEARING_BLINKER;
      O     "Timer 0";
      =     "H 52.0";
END_FUNCTION

FUNCTION "HMI CONTROL" : VOID
TITLE =HMI Control - Screen 0 SSW Inputs
//Screen 0 - "RUN" Screen
NAME : HMI_CTRL
VERSION : 0.1


VAR_TEMP
  SERVICE_ON : BOOL ;
  CLEARING_ON : BOOL ;
  HAND_FEED : BOOL ;
  UPDATE_PULSE : BOOL ;
END_VAR
BEGIN
NETWORK
TITLE =New HMI Panel Switches
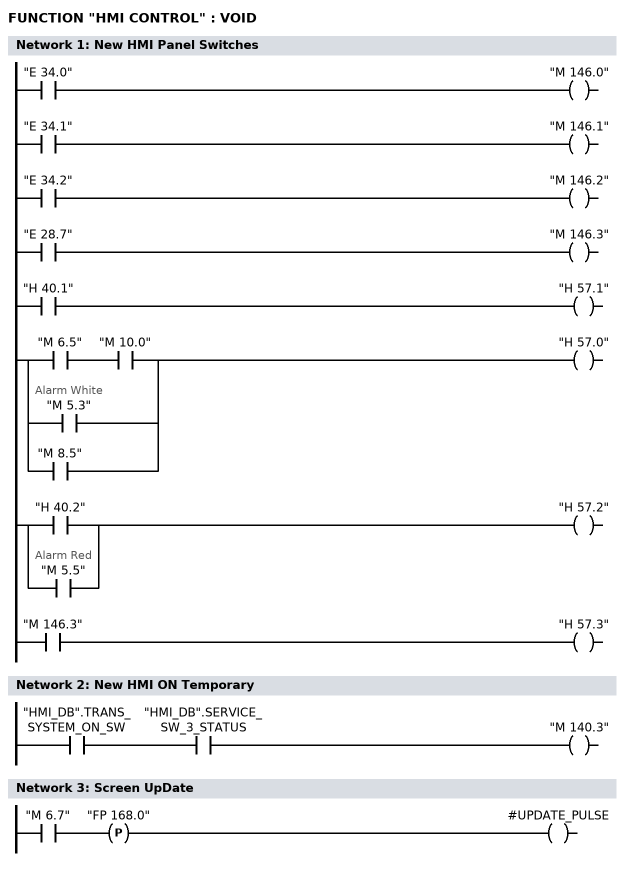

      A     "E 34.0";
      =     "M 146.0";
//;
      A     "E 34.1";
      =     "M 146.1";
//;
      A     "E 34.2";
      =     "M 146.2";
//;
      A     "E 28.7";
      =     "M 146.3";
//;
      A     "H 40.1";
      =     "H 57.1";
//;
      A(    ;
      A     "M 6.5";
      A     "M 10.0";
      )     ;
      O     "M 5.3"; // Alarm White
      O     "M 8.5";
      =     "H 57.0";
//;
      A     "H 40.2";
      O     "M 5.5"; // Alarm Red
      =     "H 57.2";
//;
      A     "M 146.3";
      =     "H 57.3";
NETWORK
TITLE =New HMI ON Temporary

      A     "HMI_DB".TRANS_SYSTEM_ON_SW;
      A     "HMI_DB".SERVICE_SW_3_STATUS;
      =     "M 140.3";
NETWORK
TITLE =Screen UpDate

      A     "M 6.7";
      FP    "FP 168.0";
      =     #UPDATE_PULSE;
NETWORK
TITLE =Screen 0 Soft Switches

      A(    ;
      L     "HMI_DB".ACTUAL_HMI_SCREEN_NO;
      L     "HMI_UPDATE".HMI_MAIN_PAGE_GRAPHIC;
      <>I   ;
      )     ;
      O     #UPDATE_PULSE;
      JNB   MAIN;
NETWORK
TITLE =Service Switch Status - Screen 0 SSW Inputs
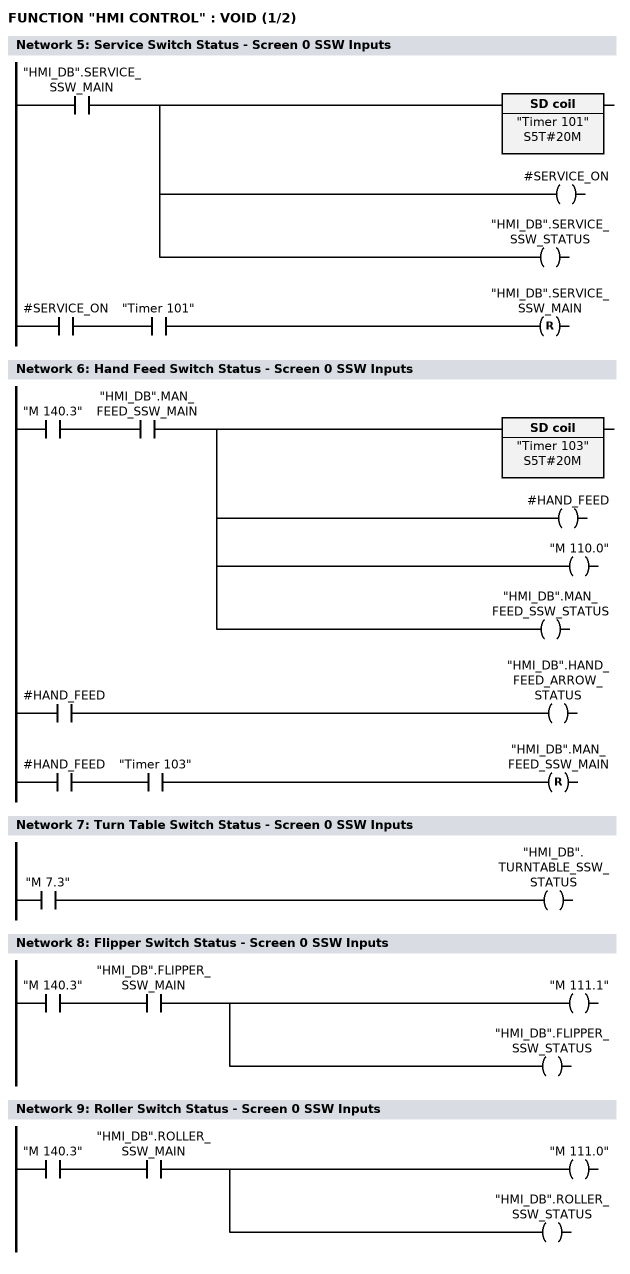

      A     "HMI_DB".SERVICE_SSW_MAIN;
      L     S5T#20M;
      SD    "Timer 101";
      =     #SERVICE_ON;
      =     "HMI_DB".SERVICE_SSW_STATUS;
//;
      A     #SERVICE_ON;
      A     "Timer 101";
      R     "HMI_DB".SERVICE_SSW_MAIN;
NETWORK
TITLE =Hand Feed Switch Status - Screen 0 SSW Inputs

      A     "M 140.3";
      A     "HMI_DB".MAN_FEED_SSW_MAIN;
      L     S5T#20M;
      SD    "Timer 103";
      =     #HAND_FEED;
      =     "M 110.0";
      =     "HMI_DB".MAN_FEED_SSW_STATUS;
//;
      A     #HAND_FEED;
      =     "HMI_DB".HAND_FEED_ARROW_STATUS;
//;
      A     #HAND_FEED;
      A     "Timer 103";
      R     "HMI_DB".MAN_FEED_SSW_MAIN;
NETWORK
TITLE =Turn Table Switch Status - Screen 0 SSW Inputs

      A     "M 7.3";
      =     "HMI_DB".TURNTABLE_SSW_STATUS;
NETWORK
TITLE =Flipper Switch Status - Screen 0 SSW Inputs

      A     "M 140.3";
      A     "HMI_DB".FLIPPER_SSW_MAIN;
      =     "M 111.1";
      =     "HMI_DB".FLIPPER_SSW_STATUS;
NETWORK
TITLE =Roller Switch Status - Screen 0 SSW Inputs

      A     "M 140.3";
      A     "HMI_DB".ROLLER_SSW_MAIN;
      =     "M 111.0";
      =     "HMI_DB".ROLLER_SSW_STATUS;
NETWORK
TITLE =HMI Service Switch Reset
//HMI Service Switch Reset when 2145 Exits Packets + 10s Delay
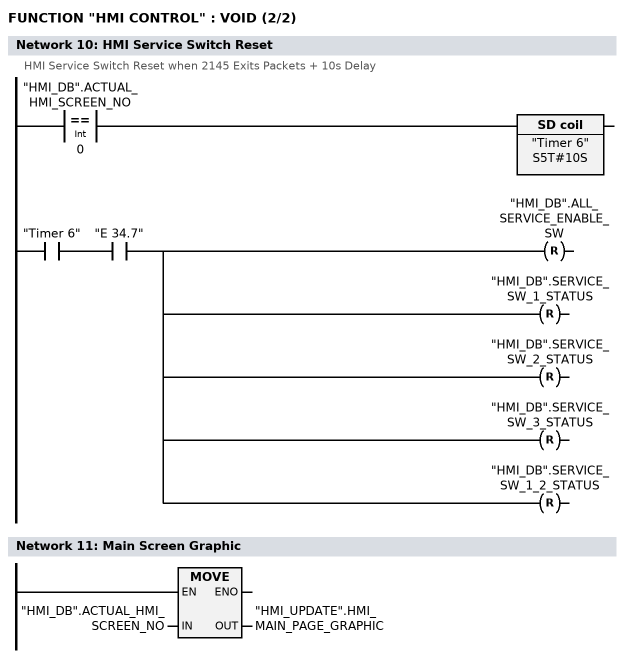
      A(    ;
      L     "HMI_DB".ACTUAL_HMI_SCREEN_NO;
      L     0;
      ==I   ;
      )     ;
      L     S5T#10S;
      SD    "Timer 6";
//;
      A     "Timer 6";
      A     "E 34.7";
      R     "HMI_DB".ALL_SERVICE_ENABLE_SW;
      R     "HMI_DB".SERVICE_SW_1_STATUS;
      R     "HMI_DB".SERVICE_SW_2_STATUS;
      R     "HMI_DB".SERVICE_SW_3_STATUS;
      R     "HMI_DB".SERVICE_SW_1_2_STATUS;
NETWORK
TITLE =Main Screen Graphic


      L     "HMI_DB".ACTUAL_HMI_SCREEN_NO;
      T     "HMI_UPDATE".HMI_MAIN_PAGE_GRAPHIC;

MAIN: NOP   0;
END_FUNCTION

FUNCTION "HMI COMMS" : VOID
TITLE =HMI Communications
//OMRON NS12  on DB12
NAME : HMI_COMM
VERSION : 0.1


VAR_TEMP
  UPDATE_PULSE_0 : BOOL ;
  UPDATE_PULSE_1 : BOOL ;
  UPDATE_PULSE_2 : BOOL ;
  UPDATE_PULSE_3 : BOOL ;
  UPDATE_PULSE_4 : BOOL ;
  UPDATE_PULSE_5 : BOOL ;
  UPDATE_PULSE_6 : BOOL ;
  UPDATE_1 : BOOL ;
  UPDATE_2 : BOOL ;
  UPDATE_3 : BOOL ;
  UPDATE_4 : BOOL ;
  UPDATE_5 : BOOL ;
  UPDATE_6 : BOOL ;
  UPDATE_7 : BOOL ;
  UPDATE_8 : BOOL ;
  UPDATE_9 : BOOL ;
  UPDATE_10 : BOOL ;
  UPDATE_11 : BOOL ;
  UPDATE_12 : BOOL ;
  UPDATE_13 : BOOL ;
  TEMP1 : BOOL ;
  TEST : BOOL ;
  CONVEYOR_0_COLOR : BYTE ;
  ELEVATOR_COLOR : BYTE ;
  CONVEYOR_1_COLOR : BYTE ;
  CONVEYOR_2_COLOR : BYTE ;
  CONVEYOR_3_COLOR : BYTE ;
  CONVEYOR_4_COLOR : BYTE ;
  CONVEYOR_5_COLOR : BYTE ;
  CONVEYOR_6_COLOR : BYTE ;
  CONVEYOR_7_COLOR : BYTE ;
  CONVEYOR_8_COLOR : BYTE ;
  CONVEYOR_9_COLOR : BYTE ;
  PUSHER_2_COLOR : BOOL ;
  CONVEYOR_11_COLOR : BYTE ;
  CONVEYOR_12_COLOR : BYTE ;
  CONVEYOR_13_COLOR : BYTE ;
  CONVEYOR_21_COLOR : BYTE ;
  CONVEYOR_22_COLOR : BYTE ;
  CONVEYOR_23_COLOR : BYTE ;
  CONVEYOR_10_COLOR : BYTE ;
  NEW_ORDER_COLOR : BYTE ;
END_VAR
BEGIN
NETWORK
TITLE =HMI - UpDate Timing
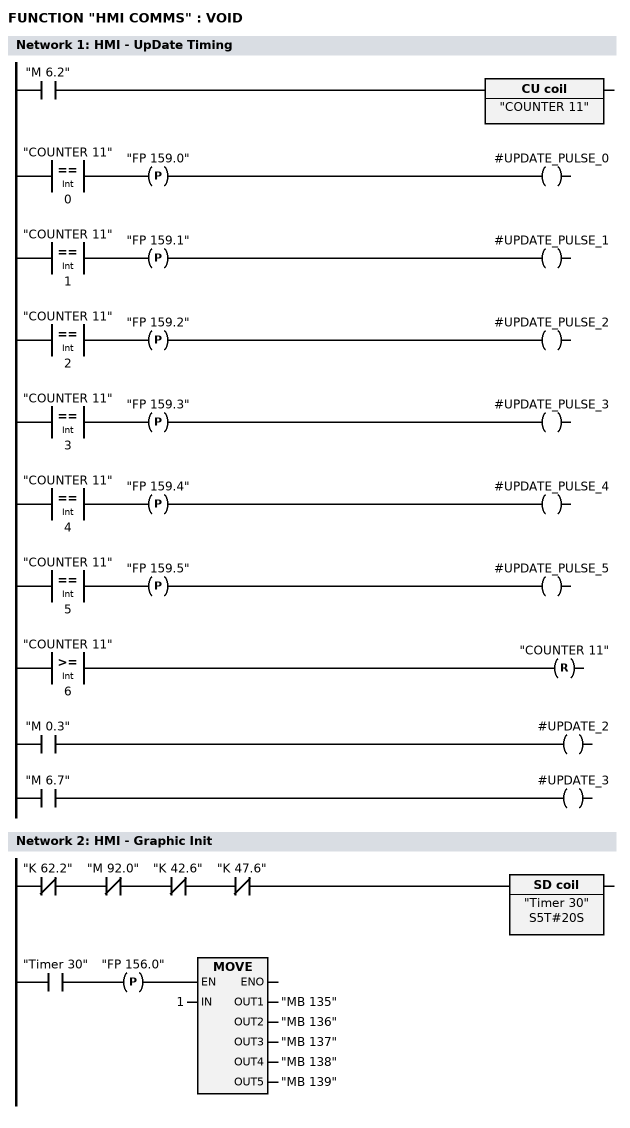

      A     "M 6.2";
      CU    "COUNTER 11";
//;
      A(    ;
      L     "COUNTER 11";
      L     0;
      ==I   ;
      )     ;
      FP    "FP 159.0";
      =     #UPDATE_PULSE_0;
//;
      A(    ;
      L     "COUNTER 11";
      L     1;
      ==I   ;
      )     ;
      FP    "FP 159.1";
      =     #UPDATE_PULSE_1;
//;
      A(    ;
      L     "COUNTER 11";
      L     2;
      ==I   ;
      )     ;
      FP    "FP 159.2";
      =     #UPDATE_PULSE_2;
//;
      A(    ;
      L     "COUNTER 11";
      L     3;
      ==I   ;
      )     ;
      FP    "FP 159.3";
      =     #UPDATE_PULSE_3;
//;
      A(    ;
      L     "COUNTER 11";
      L     4;
      ==I   ;
      )     ;
      FP    "FP 159.4";
      =     #UPDATE_PULSE_4;
//;
      A(    ;
      L     "COUNTER 11";
      L     5;
      ==I   ;
      )     ;
      FP    "FP 159.5";
      =     #UPDATE_PULSE_5;
//;
      A(    ;
      L     "COUNTER 11";
      L     6;
      >=I   ;
      )     ;
      R     "COUNTER 11";
//;;
      A     "M 0.3";
      =     #UPDATE_2;
//;
      A     "M 6.7";
      =     #UPDATE_3;
NETWORK
TITLE =HMI - Graphic Init

      AN    "K 62.2";
      AN    "M 92.0";
      AN    "K 42.6";
      AN    "K 47.6";
      L     S5T#20S;
      SD    "Timer 30";
//;
      A     "Timer 30";
      FP    "FP 156.0";
      JNB   K622;
      L     1;
      T     "MB 135";
      T     "MB 136";
      T     "MB 137";
      T     "MB 138";
      T     "MB 139";

K622: NOP   0;
NETWORK
TITLE =HMI - Doors Monitor

      ON    "E 4.6";
      ON    "E 9.0";
      ON    "E 12.5";
      O     #UPDATE_PULSE_0;
      JNB   DOOR;
      AN    "E 4.6";
      =     "HMI_DB".ELEVATOR_DOOR_STATUS;
//;
      AN    "E 9.0";
      =     "HMI_DB".FLIPPER_DOOR_STATUS;
//;
      AN    "E 12.5";
      =     "HMI_DB".LOADER_DOOR_STATUS;

DOOR: NOP   0;
NETWORK
TITLE =HMI - E-Stop Monitor

      O     "M 1.0";
      O     "M 1.1";
      O     "M 1.2";
      O     "M 1.3";
      O     #UPDATE_PULSE_1;
      JNB   ESTP;
      A     "M 1.0";
      =     "HMI_DB".E_STOP_CONSOLE_STATUS;
//;
      A     "M 1.1";
      =     "HMI_DB".E_STOP_LOADER_STATUS;
//;
      A     "M 1.2";
      =     "HMI_DB".E_STOP_ELEVATOR_STATUS;
//;
      A     "M 1.3";
      =     "HMI_DB".E_STOP_FLIPPER_STATUS;

ESTP: NOP   0;
NETWORK
TITLE =HMI - Motors Fault Status

      A(    ;
      L     "MW 2";
      L     0;
      <>I   ;
      O     ;
      L     "MB 4";
      L     0;
      <>I   ;
      )     ;
      O     "M 7.0";
      O     "M 7.1";
      O     "M 7.2";
      O     #UPDATE_PULSE_2;
      JNB   MTRF;
      A     "M 2.0";
      =     "HMI_DB".CONVEYOR_0_MOTOR_STATUS;
//;
      A     "M 2.1";
      =     "HMI_DB".PUSHER_0_MOTOR_STATUS;
//;
      A     "M 2.2";
      =     "HMI_DB".ELEVATOR_MOTOR_STATUS;
//;
      A     "M 2.3";
      =     "HMI_DB".PUSHER_1_MOTOR_STATUS;
//;
      A     "M 2.4";
      =     "HMI_DB".CONVEYOR_1_MOTOR_STATUS;
//;
      A     "M 2.5";
      =     "HMI_DB".CONVEYOR_2B_MOTOR_STATUS;
//;
      A     "M 2.6";
      =     "HMI_DB".CONVEYOR_2R_MOTOR_STATUS;
//;
      A     "M 2.7";
      =     "HMI_DB".CONVEYOR_3_MOTOR_STATUS;
//;
      A     "M 3.0";
      =     "HMI_DB".CONVEYOR_4_MOTOR_STATUS;
//;
      A     "M 3.1";
      =     "HMI_DB".CONVEYOR_5_MOTOR_STATUS;
//;
      A     "M 3.2";
      =     "HMI_DB".CONVEYOR_6_MOTOR_STATUS;
//;
      A     "M 3.3";
      =     "HMI_DB".CONVEYOR_7_MOTOR_STATUS;
//;
      A     "M 3.4";
      =     "HMI_DB".FLIPPER_MOTOR_STATUS;
//;
      A     "M 3.5";
      =     "HMI_DB".CONVEYOR_8_MOTOR_STATUS;
//;
      A     "M 3.6";
      =     "HMI_DB".TURNTABLE_MOTOR_STATUS;
//;
      A     "M 3.7";
      =     "HMI_DB".CONVEYOR_9_MOTOR_STATUS;
//;
      A     "M 4.0";
      =     "HMI_DB".PUSHER_2_MOTOR_STATUS;
//;
      A     "M 4.1";
      =     "HMI_DB".CONVEYOR_10_MOTOR_STATUS;
//;
      A     "M 4.2";
      =     "HMI_DB".CONVEYOR_11_MOTOR_STATUS;
//;
      A     "M 4.3";
      =     "HMI_DB".CONVEYOR_12_MOTOR_STATUS;
//;
      A     "M 4.4";
      =     "HMI_DB".CONVEYOR_13_MOTOR_STATUS;
//;
      A     "M 4.5";
      =     "HMI_DB".CONVEYOR_21_MOTOR_STATUS;
//;
      A     "M 4.6";
      =     "HMI_DB".CONVEYOR_22_MOTOR_STATUS;
//;
      A     "M 4.7";
      =     "HMI_DB".CONVEYOR_23_MOTOR_STATUS;
//;
      A     "M 7.0";
      =     "HMI_DB".LOADER_LIFT_MOTOR_STATUS;
//;
      A     "M 7.1";
      =     "HMI_DB".LOADER_FING_MOTOR_STATUS;
//;
      A     "M 7.2";
      =     "HMI_DB".LOADER_BELT_MOTOR_STATUS;

MTRF: NOP   0;
NETWORK
TITLE =HMI Light Barriers Status - Conveyors 1, 2, 3 LBs

      A(    ;
      L     IW     5;
      L     "HMI_UPDATE".HMI_GRAPHIC_TOTAL_1;
      <>I   ;
      O     #UPDATE_PULSE_3;
      )     ;
      JNB   LBS1;
      A     "B 5.4";
      =     "HMI_DB".LIGHT_BARRIER_1_STATUS;
//;
      A     "B 5.5";
      =     "HMI_DB".LIGHT_BARRIER_2_STATUS;
//;
      A     "B 6.0";
      =     "HMI_DB".LIGHT_BARRIER_3_STATUS;
//;
      A     "B 6.1";
      =     "HMI_DB".LIGHT_BARRIER_4_STATUS;
//;
      A     "B 6.2";
      =     "HMI_DB".LIGHT_BARRIER_5_STATUS;
//;
      A     "B 6.4";
      =     "HMI_DB".LIGHT_BARRIER_6_STATUS;
//;
      A     "B 5.2";
      =     "HMI_DB".LIGHT_BARRIER_B_STATUS;
//;
      A     "B 5.1";
      =     "HMI_DB".LIGHT_BARRIER_A_STATUS;
//;
      L     IW     5;
      T     "HMI_UPDATE".HMI_GRAPHIC_TOTAL_1;

LBS1: NOP   0;
NETWORK
TITLE =HMI Light Barriers Status - Conveyors 4, 5, 6, 7, 8, 9 LBs

      A(    ;
      L     IW     6;
      L     "HMI_UPDATE".HMI_GRAPHIC_TOTAL_2;
      <>I   ;
      O     #UPDATE_PULSE_4;
      )     ;
      O     "B 8.2";
      JNB   LBS2;
      A     "B 6.7";
      =     "HMI_DB".LIGHT_BARRIER_7_STATUS;
//;
      A     "B 7.0";
      =     "HMI_DB".LIGHT_BARRIER_8_STATUS;
//;
      A     "B 7.1";
      =     "HMI_DB".LIGHT_BARRIER_9_STATUS;
//;
      A     "B 7.2";
      =     "HMI_DB".LIGHT_BARRIER_10_STATUS;
//;
      A     "B 7.3";
      =     "HMI_DB".LIGHT_BARRIER_11_STATUS;
//;
      A     "B 7.4";
      =     "HMI_DB".LIGHT_BARRIER_12_STATUS;
//;
      A     "B 8.2";
      =     "HMI_DB".LIGHT_BARRIER_13_STATUS;
//;
      L     IW     6;
      T     "HMI_UPDATE".HMI_GRAPHIC_TOTAL_2;

LBS2: NOP   0;
NETWORK
TITLE =HMI Light Barriers Status - Conveyors 10, 11, 12, 13, 21, 22, 23

      A(    ;
      L     IW     9;
      L     IW    12;
      +I    ;
      L     IB    15;
      +I    ;
      L     "HMI_UPDATE".HMI_FEED_GRAPHIC;
      <>I   ;
      O     #UPDATE_PULSE_5;
      )     ;
      JNB   LBS3;
      A     "B 9.6";
      =     "HMI_DB".LIGHT_BARRIER_14_STATUS;
//;
      A     "B 9.7";
      =     "HMI_DB".LIGHT_BARRIER_15_STATUS;
//;
      A     "B 10.3";
      =     "HMI_DB".LIGHT_BARRIER_16_STATUS;
//;
      A     "B 10.4";
      =     "HMI_DB".LIGHT_BARRIER_17_STATUS;
//;
      A     "B 10.5";
      =     "HMI_DB".LIGHT_BARRIER_18_STATUS;
//;
      A     "B 10.6";
      =     "HMI_DB".LIGHT_BARRIER_19_STATUS;
//;
      A     "B 10.7";
      =     "HMI_DB".LIGHT_BARRIER_20_STATUS;
//;
      A     "B 11.0";
      =     "HMI_DB".LIGHT_BARRIER_21_STATUS;
//;
      A     "B 11.1";
      =     "HMI_DB".LIGHT_BARRIER_22_STATUS;
//;
      A     "B 11.2";
      =     "HMI_DB".LIGHT_BARRIER_23_STATUS;
//;
      A     "B 12.3";
      =     "HMI_DB".LIGHT_BARRIER_24_STATUS;
//;
      A     "B 13.0";
      =     "HMI_DB".LIGHT_BARRIER_25_STATUS;
//;
      A     "B 15.4";
      =     "HMI_DB".LIGHT_BARRIER_26_STATUS;
//;
      A     "B 15.5";
      =     "HMI_DB".LIGHT_BARRIER_27_STATUS;
//;
      A     "B 15.6";
      =     "HMI_DB".LIGHT_BARRIER_28_STATUS;
//;
      A     "B 15.7";
      =     "HMI_DB".LIGHT_BARRIER_29_STATUS;
//;
      L     IW     9;
      L     IW    12;
      +I    ;
      L     IB    15;
      +I    ;
      T     "HMI_UPDATE".HMI_FEED_GRAPHIC;

LBS3: NOP   0;
NETWORK
TITLE =HMI Light Barriers Status - Conveyors 0 LBs

      A(    ;
      L     QB    62;
      L     "HMI_UPDATE".HMI_MOTOR_TOTAL_1;
      <>I   ;
      O     #UPDATE_PULSE_0;
      )     ;
      O     "B 8.2";
      JNB   LBS4;
      A     "E 34.7";
      =     "HMI_DB".PACKETIZER_GATE_STATUS;
//;
      A     "B 35.2";
      =     "HMI_DB".LIGHT_BARRIER_30_STATUS;
//;
      A     "B 35.3";
      =     "HMI_DB".LIGHT_BARRIER_31_STATUS;
//;
      A     "B 35.4";
      =     "HMI_DB".LIGHT_BARRIER_32_STATUS;
//;
      L     QB    62;
      T     "HMI_UPDATE".HMI_MOTOR_TOTAL_1;

LBS4: NOP   0;
NETWORK
TITLE =HMI Prox Sensors Status - Elevator - Proxs

      A(    ;
      L     IB     4;
      L     "HMI_UPDATE".HMI_ELEVATOR_PROXS;
      <>I   ;
      O     #UPDATE_PULSE_1;
      )     ;
      JNB   PRX1;
      AN    "P 4.0";
      =     "HMI_DB".PROX_1_STATUS;
//;
      AN    "P 4.1";
      =     "HMI_DB".PROX_2_STATUS;
//;
      AN    "P 4.2";
      =     "HMI_DB".PROX_3_STATUS;
//;
      AN    "P 4.3";
      =     "HMI_DB".PROX_4_STATUS;
//;
      AN    "P 4.4";
      =     "HMI_DB".PROX_5_STATUS;
//;
      AN    "P 4.5";
      =     "HMI_DB".PROX_6_STATUS;
//;
      L     IB     4;
      T     "HMI_UPDATE".HMI_ELEVATOR_PROXS;

PRX1: NOP   0;
NETWORK
TITLE =HMI Prox Sensors Status - Flipper / TurnTable - Proxs

      A(    ;
      L     IW     8;
      L     "HMI_UPDATE".HMI_FLIPPER_PROXS;
      <>I   ;
      O     #UPDATE_PULSE_2;
      )     ;
      JNB   PRX2;
      AN    "P 8.0";
      =     "HMI_DB".PROX_8_STATUS;
//;
      AN    "P 8.1";
      =     "HMI_DB".PROX_7_STATUS;
//;
      AN    "P 8.5";
      =     "HMI_DB".PROX_9_STATUS;
//;
      AN    "P 8.6";
      =     "HMI_DB".PROX_10_STATUS;
//;
      AN    "P 9.2";
      =     "HMI_DB".PROX_11_STATUS;
//;
      AN    "P 9.3";
      =     "HMI_DB".PROX_12_STATUS;
//;
      L     IW     8;
      T     "HMI_UPDATE".HMI_FLIPPER_PROXS;

PRX2: NOP   0;
NETWORK
TITLE =HMI Prox Sensors Status - Pusher 2 / Pivot 10 - Proxs

      A(    ;
      L     IB    10;
      L     IB    15;
      +I    ;
      L     "HMI_UPDATE".HMI_PUSHER_PROXS;
      <>I   ;
      O     #UPDATE_PULSE_3;
      )     ;
      JNB   PRX3;
      AN    "P 10.0";
      =     "HMI_DB".PROX_13_STATUS;
//;
      AN    "P 10.1";
      =     "HMI_DB".PROX_14_STATUS;
//;
      A     "P 15.0";
      =     "HMI_DB".PROX_15_STATUS;
//;
      A     "P 15.1";
      =     "HMI_DB".PROX_16_STATUS;
//;
      L     IB    10;
      L     IB    15;
      +I    ;
      T     "HMI_UPDATE".HMI_PUSHER_PROXS;

PRX3: NOP   0;
NETWORK
TITLE =HMI Prox Sensors Status - Feeder - Proxs

      A(    ;
      L     IW    11;
      L     IB    13;
      +I    ;
      L     "HMI_UPDATE".HMI_FEEDER_PROXS;
      <>I   ;
      O     #UPDATE_PULSE_4;
      )     ;
      JNB   PRX4;
      AN    "P 13.2";
      =     "HMI_DB".PROX_17_STATUS;
//;
      AN    "P 13.1";
      =     "HMI_DB".PROX_18_STATUS;
//;
      AN    "P 11.4";
      =     "HMI_DB".PROX_19_STATUS;
//;
      AN    "P 11.5";
      =     "HMI_DB".PROX_20_STATUS;
//;
      AN    "P 11.6";
      =     "HMI_DB".PROX_21_STATUS;
//;
      AN    "P 11.7";
      =     "HMI_DB".PROX_22_STATUS;
//;
      A     "P 12.0";
      =     "HMI_DB".PROX_23_STATUS;
//;
      A     "P 12.1";
      =     "HMI_DB".PROX_24_STATUS;
//;
      L     IW    11;
      L     IB    13;
      +I    ;
      T     "HMI_UPDATE".HMI_FEEDER_PROXS;

PRX4: NOP   0;
NETWORK
TITLE =HMI - Pusher 0 - Graphic

      A(    ;
      O     "K 62.2";
      O     "K 62.3";
      O     #UPDATE_PULSE_5;
      )     ;
      JNB   PUS0;
      A     "K 62.2";
      AN    "K 62.3";
      A     "M 6.1";
      AN(   ;
      L     "MB 135";
      L     L#128;
      >=I   ;
      )     ;
      FP    "FP 156.1";
      JNB   E622;
      L     "MB 135";
      SLW   1;
      T     "MB 135";

E622: NOP   0;

      A     "K 62.3";
      AN    "K 62.2";
      A     "M 6.1";
      AN(   ;
      L     "MB 135";
      L     L#1;
      <=I   ;
      )     ;
      FP    "FP 156.2";
      JNB   R623;
      L     "MB 135";
      SRW   1;
      T     "MB 135";

R623: NOP   0;

      A     "M 6.1";
      FP    "HMI_DB".FP133;
      JNB   P133;
      L     L#255;
      L     "MB 135";
      -I    ;
      T     DB12.DBB    4;

P133: NOP   0;

PUS0: NOP   0;
NETWORK
TITLE =HMI - Elevator - Graphic

      A(    ;
      O     "M 92.0";
      O     "M 92.1";
      O     #UPDATE_PULSE_0;
      )     ;
      JNB   ELEV;
      A     "M 92.0";
      AN    "M 92.1";
      A     "M 6.2";
      AN(   ;
      L     "MB 136";
      L     L#128;
      >=I   ;
      )     ;
      FP    "FP 156.3";
      JNB   R420;
      L     "MB 136";
      SLW   1;
      T     "MB 136";

R420: NOP   0;

      A     "M 92.1";
      AN    "M 92.0";
      A     "M 6.2";
      AN(   ;
      L     "MB 136";
      L     L#1;
      <=I   ;
      )     ;
      FP    "FP 156.4";
      JNB   F420;
      L     "MB 136";
      SRW   1;
      T     "MB 136";

F420: NOP   0;

      A     "M 6.2";
      FP    "HMI_DB".FP134;
      JNB   P134;
      L     L#255;
      L     "MB 136";
      -I    ;
      T     DB12.DBB    5;

P134: NOP   0;

ELEV: NOP   0;
NETWORK
TITLE =HMI - Pusher 1 - Graphic

      A(    ;
      O     "K 42.6";
      O     "K 42.7";
      O     #UPDATE_PULSE_1;
      )     ;
      JNB   PUS1;
      A     "K 42.6";
      AN    "K 42.7";
      A     "M 6.1";
      AN(   ;
      L     "MB 137";
      L     L#128;
      >=I   ;
      )     ;
      FP    "FP 156.5";
      JNB   E426;
      L     "MB 137";
      SLW   1;
      T     "MB 137";

E426: NOP   0;

      A     "K 42.7";
      AN    "K 42.6";
      A     "M 6.1";
      AN(   ;
      L     "MB 137";
      L     L#1;
      <=I   ;
      )     ;
      FP    "FP 156.6";
      JNB   R427;
      L     "MB 137";
      SRW   1;
      T     "MB 137";

R427: NOP   0;

      A     "M 6.1";
      FP    "HMI_DB".FP135;
      JNB   P135;
      L     L#255;
      L     "MB 137";
      -I    ;
      T     DB12.DBB    6;

P135: NOP   0;

PUS1: NOP   0;
NETWORK
TITLE =HMI - Flipper Graphic

      A(    ;
      O     "K 46.0";
      O     "K 46.1";
      O     #UPDATE_PULSE_2;
      )     ;
      JNB   FLPN;
      L     3;
      A     "P 8.0";
      A     "P 8.1";
      JC    FLIP;
      L     0;

FLIP: T     "HMI_DB".FLIPPER_TURN_COLOR;

      L     1;
      AN    "P 8.0";
      A     "P 8.1";
      JC    CCW1;
      L     "HMI_DB".FLIPPER_TURN_COLOR;

CCW1: T     "HMI_DB".FLIPPER_CCW;

      L     1;
      AN    "P 8.1";
      A     "P 8.0";
      JC    CW1;
      L     "HMI_DB".FLIPPER_TURN_COLOR;

CW1:  T     "HMI_DB".FLIPPER_CW;

      L     6;
      A     "M 42.0";
      JC    FLON;
      L     9;

FLON: T     "HMI_DB".FLIPPER_COLOR;

FLPN: NOP   0;
NETWORK
TITLE =HMI - TurnTable Graphic

      A(    ;
      O     "A 47.0";
      O     "A 47.1";
      O     #UPDATE_PULSE_3;
      )     ;
      JNB   TURN;
      A(    ;
      ON    "P 9.2";
      ON    "P 9.3";
      )     ;
      S     "HMI_DB".TURNTABLE_DELIV_POSITION;
//;
      A(    ;
      ON    "P 8.5";
      ON    "P 8.6";
      )     ;
      R     "HMI_DB".TURNTABLE_DELIV_POSITION;
//;
      AN    "M 7.3";
      =     "HMI_DB".TURNTABLE_REVERSE_ARROW;
//;
      A     "M 7.3";
      =     "HMI_DB".TURNTABLE_DIR_SELECT_SW;

TURN: NOP   0;

NETWORK
TITLE =HMI - Pusher 2 - Graphic

      A(    ;
      O     "K 47.6";
      O     "K 47.7";
      O     #UPDATE_PULSE_4;
      )     ;
      JNB   PUS2;
      A     "K 47.6";
      AN    "K 47.7";
      A     "M 6.1";
      AN(   ;
      L     "MB 138";
      L     L#128;
      >=I   ;
      )     ;
      FP    "FP 156.7";
      JNB   E476;
      L     "MB 138";
      SLW   1;
      T     "MB 138";

E476: NOP   0;

      A     "K 47.7";
      AN    "K 47.6";
      A     "M 6.1";
      AN(   ;
      L     "MB 138";
      L     L#1;
      <=I   ;
      )     ;
      FP    "FP 157.0";
      JNB   R477;
      L     "MB 138";
      SRW   1;
      T     "MB 138";

R477: NOP   0;

      A     "M 6.1";
      FP    "HMI_DB".FP140;
      JNB   P140;
      L     L#255;
      L     "MB 138";
      -I    ;
      T     DB12.DBB    7;

P140: NOP   0;

PUS2: NOP   0;
NETWORK
TITLE =HMI - Pivot Graphic

      A(    ;
      O     "K 53.0";
      O     "K 53.1";
      O     #UPDATE_PULSE_5;
      )     ;
      JNB   PIVO;
      AN    "P 15.1";
      =     DB12.DBX   88.1;
//;
      AN    "P 15.0";
      =     DB12.DBX   88.0;
//;
      AN    "P 15.0";
      AN    "P 15.1";
      =     DB12.DBX   88.2;

PIVO: NOP   0;
NETWORK
TITLE =HMI - Feeder Graphic

      A(    ;
      L     IW    11;
      L     IB    13;
      +I    ;
      L     "HMI_UPDATE".HMI_FEEDER_GRAPHIC;
      <>I   ;
      O     #UPDATE_PULSE_0;
      )     ;
      JNB   FEED;

      A     "P 13.2";
      AN    "P 11.4";
      O     ;
      A     "P 11.5";
      AN    "P 11.4";
      JNB   M131;
      L     L#64;
      T     "MB 139";

M131: NOP   0;

      AN    "P 13.2";
      AN    "P 13.1";
      AN    "P 11.4";
      JNB   M132;
      L     L#128;
      T     "MB 139";

M132: NOP   0;

      AN    "P 11.4";
      AN    "P 11.5";
      JNB   M114;
      L     L#32;
      T     "MB 139";

M114: NOP   0;

      A     "P 11.4";
      AN    "P 11.5";
      A     "A 50.1";
      S     "M 70.5";
//;
      A(    ;
      A     "M 70.6";
      A     "A 50.0";
      AN    "P 11.5";
      O     ;
      A     "M 70.5";
      A     "A 50.1";
      )     ;
      JNB   M115;
      L     L#16;
      T     "MB 139";
      R     "M 70.6";

M115: NOP   0;

      A     "P 11.7";
      AN    "P 11.6";
      A     "A 50.0";
      S     "M 70.6";
//;
      A(    ;
      A     "M 70.5";
      A     "A 50.1";
      AN    "P 11.6";
      O     ;
      A     "M 70.6";
      A     "A 50.0";
      )     ;
      JNB   M116;
      L     L#8;
      T     "MB 139";
      R     "M 70.5";

M116: NOP   0;

      AN    "E 12.2";
      AN    "P 11.7";
      AN    "P 12.1";
      JNB   M117;
      L     L#4;
      T     "MB 139";

M117: NOP   0;

      AN    "E 12.2";
      AN    "P 11.7";
      A     "P 12.1";
      JNB   M121;
      L     L#6;
      T     "MB 139";

M121: NOP   0;

      A     "E 12.2";
      AN    "P 11.7";
      A     "P 12.1";
      JNB   M122;
      L     L#1;
      T     "MB 139";

M122: NOP   0;

      A     "M 6.2";
      FP    "HMI_DB".FP141;
      JNB   P141;
      L     L#255;
      L     "MB 139";
      -I    ;
      T     DB12.DBB   19;

P141: NOP   0;

      L     IW    11;
      L     IB    13;
      +I    ;
      T     "HMI_UPDATE".HMI_FEEDER_GRAPHIC;

FEED: NOP   0;
NETWORK
TITLE =HMI - Motor Run Status

      A(    ;
      L     QW    42;
      L     QW    44;
      +I    ;
      L     QW    46;
      +I    ;
      L     QW    48;
      +I    ;
      L     QW    50;
      +I    ;
      L     QB    53;
      +I    ;
      L     QB    54;
      +I    ;
      L     "HMI_UPDATE".HMI_MOTOR_GRAPHIC;
      <>I   ;
      O     #UPDATE_PULSE_1;
      )     ;
      JNB   MTR;
      O     "K 62.0";
      O     "K 62.1";
      L     0;
      JCN   K620;
      A     "K 62.0";
      L     3;
      JC    K620;
      L     6;
K620: T     "HMI_DB".CONV_0_COLOR_WORD;

      L     5;
      A     "M 14.7";
      O     "M 100.2";
      JC    E00;
      L     0;
E00:  T     #ELEVATOR_COLOR;

      L     #ELEVATOR_COLOR;
      O     "M 92.0";
      O     "M 92.1";
      JCN   Q420;
      A     "M 92.0";
      L     3;
      JC    Q420;
      L     6;
Q420: T     "HMI_DB".ELEVATOR_COLOR_WORD;

      L     0;
      A(    ;
      O     "K 42.6";
      O     "K 42.7";
      )     ;
      JCN   Q427;
      L     3;
Q427: T     "HMI_DB".PUSHER_1_COLOR_WORD;

      L     0;
      A     "A 43.0";
      JCN   Q430;
      L     3;
Q430: T     "HMI_DB".CONV_1_COLOR_WORD;

      L     5;
      A     "M 22.7";
      O     "M 100.5";
      JC    C02;
      L     0;
C02:  T     #CONVEYOR_2_COLOR;

      L     #CONVEYOR_2_COLOR;
      A     "K 43.4";
      JCN   Q434;
      L     3;
Q434: T     "HMI_DB".CONV_2_BELT_COLOR_WORD;

      L     0;
      A     "Y 43.6";
      JCN   Q436;
      L     3;
Q436: T     "HMI_DB".LIFT_ROLLER_2_COLOR_WORD;

      L     0;
      A     "K 43.5";
      JCN   Q435;
      L     3;
Q435: T     "HMI_DB".CONV_2_ROLLER_COLOR_WORD;

      L     0;
      A     "A 44.0";
      JCN   Q440;
      L     3;
Q440: T     "HMI_DB".CONV_3_COLOR_WORD;

      L     5;
      A     "M 30.7";
      O     "M 102.0";
      JC    C04;
      L     0;
C04:  T     #CONVEYOR_4_COLOR;

      L     #CONVEYOR_4_COLOR;
      A     "A 44.3";
      AN    "M 31.5";
      JCN   Q443;
      L     6;
Q443: T     "HMI_DB".CONV_4_COLOR_WORD;

      A     "A 44.3";
      A     "M 31.5";
      JNB   M315;
      L     3;
      T     "HMI_DB".CONV_4_COLOR_WORD;

M315: NOP   0;

      L     0;
      A     "A 45.0";
      JCN   Q450;
      L     3;
Q450: T     "HMI_DB".CONV_5_COLOR_WORD;

      L     5;
      A     "M 38.7";
      O     "M 102.2";
      JC    C06;
      L     0;
C06:  T     #CONVEYOR_6_COLOR;

      L     #CONVEYOR_6_COLOR;
      A     "A 45.3";
      JCN   Q453;
      L     3;
Q453: T     "HMI_DB".CONV_6_COLOR_WORD;

      L     5;
      A     "M 42.7";
      O     "M 102.3";
      JC    C07;
      L     0;
C07:  T     #CONVEYOR_7_COLOR;

      L     #CONVEYOR_7_COLOR;
      A     "A 45.6";
      JCN   Q456;
      L     3;
Q456: T     "HMI_DB".CONV_7_COLOR_WORD;

      L     0;
      A(    ;
      O     "K 46.0";
      O     "K 46.1";
      )     ;
      JCN   Q461;
      L     3;
Q461: T     "HMI_DB".FLIPPER_COLOR_WORD;

      L     0;
      A(    ;
      O     "A 47.0";
      O     "A 47.1";
      )     ;
      JCN   A470;
      L     7;

A470: T     "HMI_DB".TURN_COLOR;

//      L     0
//      AN    "M 6.2"
//      A(
//      O     "A 47.0"
//      O     "A 47.1"
//      )
//      JCN   A471
//      L     7

//A471: T     "HMI_DB".HMI_TURN_COLOR

      L     "HMI_DB".TURN_COLOR;
      A(    ;
      O     "A 46.4";
      O     "A 46.5";
      )     ;
      JCN   Q464;
      L     3;
Q464: T     "HMI_DB".CONV_8_COLOR_WORD;

      L     0;
      A     "A 47.0";
      JCN   Q470;
      L     3;
Q470: T     "HMI_DB".TURN_TABLE_COLOR_WORD;

      L     0;
      A     "K 47.5";
      JCN   Q475;
      L     3;
Q475: T     "HMI_DB".CONV_9_COLOR_WORD;

      L     0;
      A(    ;
      O     "K 47.6";
      O     "K 47.7";
      )     ;
      JCN   Q477;
      L     3;
Q477: T     "HMI_DB".PUSHER_2_COLOR_WORD;

      L     5;
      A     "M 98.1";
      O     "M 98.2";
      O     "M 106.1";
      JC    C10;
//;
      L     4;
      A     "M 55.4";
      A     "M 8.4";
      A     "M 6.5";
      JC    C10;
      L     0;

C10:  T     #CONVEYOR_10_COLOR;

      L     #CONVEYOR_10_COLOR;
      A     "A 48.0";
      A(    ;
      ON    "M 55.5";
      ON    "M 10.0";
      )     ;
      JCN   Q480;
      L     6;
Q480: T     "HMI_DB".CONV_10_COLOR_WORD;

      A     "A 48.0";
      A(    ;
      O     "M 55.5";
      O     "M 10.0";
      )     ;
      JNB   M555;
      L     3;
      T     "HMI_DB".CONV_10_COLOR_WORD;

M555: NOP   0;


      L     0;
      A     "A 48.3";
      JCN   Q483;
      L     3;
Q483: T     "HMI_DB".CONV_11_COLOR_WORD;

      L     0;
      A     "A 48.6";
      JCN   Q486;
      L     3;
Q486: T     "HMI_DB".CONV_12_COLOR_WORD;

      L     5;
      A     "M 66.7";
      O     "M 106.4";
      JC    C13;
      L     0;
C13:  T     #CONVEYOR_13_COLOR;

      L     #CONVEYOR_13_COLOR;
      A     "A 49.0";
      JCN   Q490;
      L     3;
Q490: T     "HMI_DB".CONV_13_COLOR_WORD;

      L     0;
      A     "A 53.4";
      JCN   Q534;
      L     3;
Q534: T     "HMI_DB".CONV_21_COLOR_WORD;

      L     0;
      A     "A 53.6";
      JCN   Q536;
      L     3;
Q536: T     "HMI_DB".CONV_22_COLOR_WORD;

      L     5;
      A     "M 86.7";
      O     "M 106.7";
      JC    C23;
      L     0;
C23:  T     #CONVEYOR_23_COLOR;

      L     #CONVEYOR_23_COLOR;
      A     "A 54.0";
      JCN   Q540;
      L     3;
Q540: T     "HMI_DB".CONV_23_COLOR_WORD;

      A     "M 0.7";
      =     "HMI_DB".COMPRESSED_AIR;
//;
      O     "A 50.0";
      O     "A 50.1";
      L     0;
      JCN   Q500;
      A     "A 50.0";
      L     3;
      JC    Q500;
      L     6;
Q500: T     "HMI_DB".LOADER_LIFT_COLOR_WORD;

      L     0;
      A     "A 51.0";
      JCN   Q510;
      L     3;
Q510: T     "HMI_DB".FINGERS_BELT_COLOR_WORD;

      L     QW    42;
      L     QW    44;
      +I    ;
      L     QW    46;
      +I    ;
      L     QW    48;
      +I    ;
      L     QW    50;
      +I    ;
      L     QB    53;
      +I    ;
      L     QB    54;
      +I    ;
      T     "HMI_UPDATE".HMI_MOTOR_GRAPHIC;

MTR:  NOP   0;
END_FUNCTION

FUNCTION "HMI PACKET COUNTER  NEW" : VOID
TITLE =HMI Conveyors Display Packet Counter  FC1208
//Counts are kept in "HMI_DB" (read by HMI, LIGHT BAR, C5 Re-Sync)
//Bit_0 = InFeed  /  Bit_1 = RAW Exit Sensor  /
//Transfer_Start = Transfer Step Active.
//v1.0 2026-11-23 (replaces v0.12): C11/C12/C13 + C21/C22/C23 (identical) use the
//CLEANED SENSOR LEVEL = Raw Sensor OR Blanking Active ("BLANKING DB" T_ms <
//Blank_Pct of Width_ms since the last counted front). A U-Shape sag inside the
//blanking keeps the signal ON (one packet), and a packet already ON the sensor
//when the filling step starts is still counted (v0.12 used a 400 mS pulse that
//could come before the step = first packet of a load not counted).
//FC8 settings back as v0.8 (600 / 300). Butted packets (count down): every
//"BLANKING DB".Width_ms + Gap (was #DIM_31).
//C13/C23 Count Down (once per delivery, v0.8) and C3..C10 unchanged.
//Also: duplicate presence T lines removed (no effect).
VERSION : 1.0


VAR_TEMP
  ERROR : BOOL ;
  BIT0 : BOOL ;	//Count UP Input
  XFER : BOOL ;	//Transfer Active
  BIT1 : BOOL ;	//C13/C23 Count Down Pulse - One per Delivery
  DIM_31 : INT ;	//C10 Width @ 31.0 m/min [mS]
  DIM_237 : INT ;	//C10 Width @ 23.7 m/min [mS]
  BLANK : DINT ;	//Blanking Time [mS] = Width_ms x Blank_Pct / 100
  S106 : BOOL ;	//Cleaned B10.6 - C10 Exit
  S107 : BOOL ;	//Cleaned B10.7 - C11 Exit
  S110 : BOOL ;	//Cleaned B11.0 - C12 Exit
  S154 : BOOL ;	//Cleaned B15.4 - C21 Exit
  S155 : BOOL ;	//Cleaned B15.5 - C22 Exit
END_VAR
BEGIN
NETWORK
TITLE =Packet Length mm - To Conveyor 4 HMI (as FC1206)

      L     "COLLATORS DB".PacketLength_C4;
      ITD   ;
      DTR   ;
      L     6.673000e+000;
      *R    ;
      RND   ;
      T     "MW 202";
NETWORK
TITLE =C10 Packet Width [mS] - Scaled to Link & Delivery Speeds

      L     "COLLATORS DB".Packet_Width_C10_mS; // Measured @ 27.0 m/min
      L     L#27;
      *D    ;
      L     L#31;
      /D    ;
      T     #DIM_31; // @ 31.0 m/min
//;
      L     "COLLATORS DB".Packet_Width_C10_mS;
      L     L#270;
      *D    ;
      L     L#237;
      /D    ;
      T     #DIM_237; // @ 23.7 m/min
NETWORK
TITLE =Packet Counter - Slat Conveyor 3

      A     "A 44.0";
      L     S5T#1S;
      SF    T    118; // Call Hold 1s
//;
      A     T    118;
      JNB   M440;

      L     "HMI_DB".CONVEYOR_MAXCOUNT_L;
      T     "DEBOUNCER COUNTER DB".Conveyor_C3_Slat.Maximum_Count;
      A     "B 6.2";
      =     #BIT0;
//;
      A     "A 44.0";
      =     #XFER;
//;
      CALL "DE-BOUNCER / COUNTER" (
           Bit_0                    := #BIT0,
           Bit_1                    := "B 6.4",
           Transfer_Start           := #XFER,
           Error_Reset              := "M 9.1",
           Space_DX_mS              := 600,
           ReSample_DX              := 85,
           Conveyor_Type            := 1,
           Preset_MIN_mS            := 500,
           LowSpd_Dimension_mS      := 0,
           HighSpd_Dimension_mS     := 0,
           Plc_Scan_mS              := "DB UTILITY".Scan_Cycle_Previous,
           Q_Error                  := #ERROR,
           Word_Count               := "HMI_DB".CONV_3_COUNT,
           IO_DB                    := "DEBOUNCER COUNTER DB".Conveyor_C3_Slat);

M440: NOP   0;
NETWORK
TITLE =Packet Counter - Collator Conveyor 4

      A     "A 44.3";
      L     S5T#1S;
      SF    T    119; // Call Hold 1s
//;
      A     T    119;
      JNB   M443;

      L     "HMI_DB".CONVEYOR_MAXCOUNT_L;
      T     "DEBOUNCER COUNTER DB".Conveyor_C4_Collator.Maximum_Count;
      A     "B 6.7";
      =     #BIT0;
//;
      A     "M 31.6";
      AN    "M 31.7";
      =     #XFER;
//;
      CALL "DE-BOUNCER / COUNTER" (
           Bit_0                    := #BIT0,
           Bit_1                    := "B 7.0",
           Transfer_Start           := #XFER,
           Error_Reset              := "M 9.1",
           Space_DX_mS              := 600,
           ReSample_DX              := 85,
           Conveyor_Type            := 1,
           Preset_MIN_mS            := 500,
           LowSpd_Dimension_mS      := 0,
           HighSpd_Dimension_mS     := "HOUSE_KEEPING DB".C4_Packet_Length_mS,
           Plc_Scan_mS              := "DB UTILITY".Scan_Cycle_Previous,
           Q_Error                  := #ERROR,
           Word_Count               := "HMI_DB".CONV_4_COUNT,
           IO_DB                    := "DEBOUNCER COUNTER DB".Conveyor_C4_Collator);

M443: NOP   0;
NETWORK
TITLE =Packet Counter - Link Conveyor 5

      A     "A 45.0";
      L     S5T#1S;
      SF    "Timer 120"; // Call Hold 1s
//;
      A     "Timer 120";
      =     "M 143.0";
      JNB   M450;

      L     "HMI_DB".CONVEYOR_MAXCOUNT_L;
      T     "DEBOUNCER COUNTER DB".Conveyor_C5_Link.Maximum_Count;
      A     "B 7.0";
      A     "M 35.1";
      AN    "M 35.2";
      =     #BIT0;
//;
      A     "M 35.3";
      AN    "M 35.4";
      =     #XFER;
//;
      CALL "DE-BOUNCER / COUNTER" (
           Bit_0                    := #BIT0,
           Bit_1                    := "B 7.1",
           Transfer_Start           := #XFER,
           Error_Reset              := "M 9.1",
           Space_DX_mS              := 600,
           ReSample_DX              := 85,
           Conveyor_Type            := 3,
           Preset_MIN_mS            := 500,
           LowSpd_Dimension_mS      := 0,
           HighSpd_Dimension_mS     := "HOUSE_KEEPING DB".C4_Packet_Length_mS,
           Plc_Scan_mS              := "DB UTILITY".Scan_Cycle_Previous,
           Q_Error                  := #ERROR,
           Word_Count               := "HMI_DB".CONV_5_COUNT,
           IO_DB                    := "DEBOUNCER COUNTER DB".Conveyor_C5_Link);

M450: NOP   0;
NETWORK
TITLE =Packet Counter - Delivery Conveyor 6

      A     "A 45.3";
      L     S5T#1S;
      SF    "Timer 121"; // Call Hold 1s
//;
      A     "Timer 121";
      =     "M 143.1";
      JNB   M453;

      L     "HMI_DB".CONVEYOR_MAXCOUNT_L;
      T     "DEBOUNCER COUNTER DB".Conveyor_C6_Delivery.Maximum_Count;
      A     "B 7.1";
      A     "M 39.1";
      AN    "M 39.2";
      =     #BIT0;
//;
      A     "M 39.4";
      AN    "M 39.5";
      =     #XFER;
//;
      CALL "DE-BOUNCER / COUNTER" (
           Bit_0                    := #BIT0,
           Bit_1                    := "B 7.3",
           Transfer_Start           := #XFER,
           Error_Reset              := "M 9.1",
           Space_DX_mS              := 600,
           ReSample_DX              := 85,
           Conveyor_Type            := 2,
           Preset_MIN_mS            := 500,
           LowSpd_Dimension_mS      := 0,
           HighSpd_Dimension_mS     := "HOUSE_KEEPING DB".C4_Packet_Length_mS,
           Plc_Scan_mS              := "DB UTILITY".Scan_Cycle_Previous,
           Q_Error                  := #ERROR,
           Word_Count               := "HMI_DB".CONV_6_COUNT,
           IO_DB                    := "DEBOUNCER COUNTER DB".Conveyor_C6_Delivery);

M453: NOP   0;
NETWORK
TITLE =Packet Presence - Flipper / TurnTable / Conveyor 9 / Pusher 2

      L     0;
      A     "M 43.4";
      JCN   M434;

      L     1;

M434: T     "HMI_DB".FLIPPER_PACK_PRESENCE;
//;
      L     0;
      A     "M 47.4";
      JCN   M474;

      L     1;

M474: T     "HMI_DB".TURNTABLE_PACK_PRESENCE;
//;
      L     0;
      A     "M 51.4";
      JCN   M514;

      L     1;

M514: T     "HMI_DB".ROLLER_PACK_PRESENCE;
//;
      L     0;
      A     "M 51.5";
      JCN   M515;

      L     1;

M515: T     "HMI_DB".PUSHER_PACK_PRESENCE;
NETWORK
TITLE =Packet Counter - Pivot Conveyor 10

      A     "A 48.0";
      L     S5T#1S;
      SF    T    134; // Call Hold 1s
//;
      A     T    134;
      JNB   M480;

      L     "HMI_DB".CONVEYOR_MAXCOUNT_W;
      T     "DEBOUNCER COUNTER DB".Conveyor_C10_Collator.Maximum_Count;
      A     "B 10.4";
      =     #BIT0;
//;
      A     "M 55.5";
      AN    "M 55.6";
      =     #XFER;
//;
      CALL "DE-BOUNCER / COUNTER" (
           Bit_0                    := #BIT0,
           Bit_1                    := "B 10.6",
           Transfer_Start           := #XFER,
           Error_Reset              := "M 9.1",
           Space_DX_mS              := 600,
           ReSample_DX              := 85,
           Conveyor_Type            := 1,
           Preset_MIN_mS            := 500,
           LowSpd_Dimension_mS      := 0,
           HighSpd_Dimension_mS     := #DIM_31,
           Plc_Scan_mS              := "DB UTILITY".Scan_Cycle_Previous,
           Q_Error                  := #ERROR,
           Word_Count               := "HMI_DB".CONV_10_COUNT,
           IO_DB                    := "DEBOUNCER COUNTER DB".Conveyor_C10_Collator);

M480: NOP   0;
NETWORK
TITLE =Cleaned Sensors - Raw OR Blanking Active (U-Shape Sag Filled)
//Blanking from "BLANKING DB" (FC1212 in FC1210): T_ms = belt run time since the
//last counted front at this sensor. While T_ms < Blank_Pct of the packet time
//the signal stays ON, so a sag inside a packet is not a gap.
      L     "BLANKING DB".Width_ms;
      ITD   ;
      L     "BLANKING DB".Blank_Pct;
      ITD   ;
      *D    ;
      L     L#100;
      /D    ;
      T     #BLANK;
//;
      A(    ;
      L     "BLANKING DB".C10_Exit_B10_6.T_ms;
      L     #BLANK;
      <D    ;
      )     ;
      O     "B 10.6"; // C10 Exit Sens
      =     #S106;
//;
      A(    ;
      L     "BLANKING DB".C11_Exit_B10_7.T_ms;
      L     #BLANK;
      <D    ;
      )     ;
      O     "B 10.7"; // C11 Exit Sens
      =     #S107;
//;
      A(    ;
      L     "BLANKING DB".C12_Exit_B11_0.T_ms;
      L     #BLANK;
      <D    ;
      )     ;
      O     "B 11.0"; // C12 Exit Sens
      =     #S110;
//;
      A(    ;
      L     "BLANKING DB".C21_Exit_B15_4.T_ms;
      L     #BLANK;
      <D    ;
      )     ;
      O     "B 15.4"; // C21 Exit Sens
      =     #S154;
//;
      A(    ;
      L     "BLANKING DB".C22_Exit_B15_5.T_ms;
      L     #BLANK;
      <D    ;
      )     ;
      O     "B 15.5"; // C22 Exit Sens
      =     #S155;
NETWORK
TITLE =Packet Counter - Link Conveyor 11 (Low)

      A     "A 48.3";
      L     S5T#1S;
      SF    "Timer 122"; // Call Hold 1s
//;
      A     "Timer 122";
      =     "M 143.2";
      JNB   M483;

      L     "HMI_DB".CONVEYOR_MAXCOUNT_W;
      T     "DEBOUNCER COUNTER DB".Conveyor_C11_Link.Maximum_Count;
      A     #S106; // Cleaned B 10.6
      A     "M 59.1";
      AN    "M 59.2";
      A     "P 15.1";
      =     #BIT0;
//;
      A     "M 59.3";
      AN    "M 59.4";
      =     #XFER;
//;
      CALL "DE-BOUNCER / COUNTER" (
           Bit_0                    := #BIT0,
           Bit_1                    := #S107,
           Transfer_Start           := #XFER,
           Error_Reset              := "M 9.1",
           Space_DX_mS              := 600,
           ReSample_DX              := 85,
           Conveyor_Type            := 3,
           Preset_MIN_mS            := 300,
           LowSpd_Dimension_mS      := 0,
           HighSpd_Dimension_mS     := "BLANKING DB".Width_ms,
           Plc_Scan_mS              := "DB UTILITY".Scan_Cycle_Previous,
           Q_Error                  := #ERROR,
           Word_Count               := "HMI_DB".CONV_11_COUNT,
           IO_DB                    := "DEBOUNCER COUNTER DB".Conveyor_C11_Link);

M483: NOP   0;
NETWORK
TITLE =Packet Counter - Link Conveyor 12 (Low)

      A     "A 48.6";
      L     S5T#1S;
      SF    "Timer 123"; // Call Hold 1s
//;
      A     "Timer 123";
      =     "M 143.3";
      JNB   M486;

      L     "HMI_DB".CONVEYOR_MAXCOUNT_W;
      T     "DEBOUNCER COUNTER DB".Conveyor_C12_Link.Maximum_Count;
      A     #S107; // Cleaned B 10.7
      A     "M 63.1";
      AN    "M 63.2";
      =     #BIT0;
//;
      A     "M 63.3";
      AN    "M 63.4";
      =     #XFER;
//;
      CALL "DE-BOUNCER / COUNTER" (
           Bit_0                    := #BIT0,
           Bit_1                    := #S110,
           Transfer_Start           := #XFER,
           Error_Reset              := "M 9.1",
           Space_DX_mS              := 600,
           ReSample_DX              := 85,
           Conveyor_Type            := 3,
           Preset_MIN_mS            := 300,
           LowSpd_Dimension_mS      := 0,
           HighSpd_Dimension_mS     := "BLANKING DB".Width_ms,
           Plc_Scan_mS              := "DB UTILITY".Scan_Cycle_Previous,
           Q_Error                  := #ERROR,
           Word_Count               := "HMI_DB".CONV_12_COUNT,
           IO_DB                    := "DEBOUNCER COUNTER DB".Conveyor_C12_Link);

M486: NOP   0;
NETWORK
TITLE =Packet Counter - Delivery Conveyor 13 (Low)

      A     "A 49.0";
      L     S5T#1S;
      SF    "Timer 124"; // Call Hold 1s
//;
      A     "Timer 124";
      =     "M 143.4";
      JNB   M490;

      L     "HMI_DB".CONVEYOR_MAXCOUNT_W;
      T     "DEBOUNCER COUNTER DB".Conveyor_C13_Delivery.Maximum_Count;
      A     #S110; // Cleaned B 11.0
      A     "M 67.1";
      AN    "M 67.2";
      =     #BIT0;
//;
//C13: Count Down only a packet the Exit Sens has SEEN on the edge and SEEN
//leave (Delivery Done M67.5 = B11.2 clear). Once per delivery: the sag of a
//U-Shape packet (beam at top of stack) can not count it twice.
      A     "M 67.4"; // Delivery
      AN    "M 67.5";
      A     "B 11.2"; // Packet on the Edge - Seen by Exit Sens
      S     "M 283.3"; // Packet Seen (Free)
//;
      A     "M 67.5"; // Delivery Done - Exit Sens Clear
      FP    M    283.2; // Edge Memory (Free)
      A     "M 283.3"; // Only if a Packet was Seen
      L     S5T#500MS;
      SE    "Timer 139"; // Count Down Pulse 500mS (> Preset_MIN 300mS)
//;
      A     "Timer 139"; // Counted
      O     "M 67.6"; // Steps Reset
      R     "M 283.3";
//;
      A     "Timer 139";
      =     #BIT1; // Count Down Pulse
      =     #XFER;
//;
      CALL "DE-BOUNCER / COUNTER" (
           Bit_0                    := #BIT0,
           Bit_1                    := #BIT1,
           Transfer_Start           := #XFER,
           Error_Reset              := "M 9.1",
           Space_DX_mS              := 600,
           ReSample_DX              := 85,
           Conveyor_Type            := 2,
           Preset_MIN_mS            := 300,
           LowSpd_Dimension_mS      := 0,
           HighSpd_Dimension_mS     := 0,
           Plc_Scan_mS              := "DB UTILITY".Scan_Cycle_Previous,
           Q_Error                  := #ERROR,
           Word_Count               := "HMI_DB".CONV_13_COUNT,
           IO_DB                    := "DEBOUNCER COUNTER DB".Conveyor_C13_Delivery);

M490: NOP   0;
NETWORK
TITLE =Packet Counter - Link Conveyor 21 (High)

      A     "A 53.4";
      L     S5T#1S;
      SF    "Timer 125"; // Call Hold 1s
//;
      A     "Timer 125";
      =     "M 143.5";
      JNB   M534;

      L     "HMI_DB".CONVEYOR_MAXCOUNT_W;
      T     "DEBOUNCER COUNTER DB".Conveyor_C21_Link.Maximum_Count;
      A     #S106; // Cleaned B 10.6
      A     "M 79.1";
      AN    "M 79.2";
      A     "P 15.0";
      =     #BIT0;
//;
      A     "M 79.3";
      AN    "M 79.4";
      =     #XFER;
//;
      CALL "DE-BOUNCER / COUNTER" (
           Bit_0                    := #BIT0,
           Bit_1                    := #S154,
           Transfer_Start           := #XFER,
           Error_Reset              := "M 9.1",
           Space_DX_mS              := 600,
           ReSample_DX              := 85,
           Conveyor_Type            := 3,
           Preset_MIN_mS            := 300,
           LowSpd_Dimension_mS      := 0,
           HighSpd_Dimension_mS     := "BLANKING DB".Width_ms,
           Plc_Scan_mS              := "DB UTILITY".Scan_Cycle_Previous,
           Q_Error                  := #ERROR,
           Word_Count               := "HMI_DB".CONV_21_COUNT,
           IO_DB                    := "DEBOUNCER COUNTER DB".Conveyor_C21_Link);

M534: NOP   0;
NETWORK
TITLE =Packet Counter - Link Conveyor 22 (High)

      A     "A 53.6";
      L     S5T#1S;
      SF    "Timer 126"; // Call Hold 1s
//;
      A     "Timer 126";
      =     "M 143.6";
      JNB   M536;

      L     "HMI_DB".CONVEYOR_MAXCOUNT_W;
      T     "DEBOUNCER COUNTER DB".Conveyor_C22_Link.Maximum_Count;
      A     #S154; // Cleaned B 15.4
      A     "M 83.1";
      AN    "M 83.2";
      =     #BIT0;
//;
      A     "M 83.3";
      AN    "M 83.4";
      =     #XFER;
//;
      CALL "DE-BOUNCER / COUNTER" (
           Bit_0                    := #BIT0,
           Bit_1                    := #S155,
           Transfer_Start           := #XFER,
           Error_Reset              := "M 9.1",
           Space_DX_mS              := 600,
           ReSample_DX              := 85,
           Conveyor_Type            := 3,
           Preset_MIN_mS            := 300,
           LowSpd_Dimension_mS      := 0,
           HighSpd_Dimension_mS     := "BLANKING DB".Width_ms,
           Plc_Scan_mS              := "DB UTILITY".Scan_Cycle_Previous,
           Q_Error                  := #ERROR,
           Word_Count               := "HMI_DB".CONV_22_COUNT,
           IO_DB                    := "DEBOUNCER COUNTER DB".Conveyor_C22_Link);

M536: NOP   0;
NETWORK
TITLE =Packet Counter - Delivery Conveyor 23 (High)

      A     "A 54.0";
      L     S5T#1S;
      SF    "Timer 127"; // Call Hold 1s
//;
      A     "Timer 127";
      =     "M 143.7";
      JNB   M540;

      L     "HMI_DB".CONVEYOR_MAXCOUNT_W;
      T     "DEBOUNCER COUNTER DB".Conveyor_C23_Delivery.Maximum_Count;
      A     #S155; // Cleaned B 15.5
      A     "M 87.1";
      AN    "M 87.2";
      =     #BIT0;
//;
//C23: Count Down only a packet the Exit Sens has SEEN on the edge and SEEN
//leave (Delivery Done M87.5 = B15.7 clear). Once per delivery: the sag of a
//U-Shape packet (beam at top of stack) can not count it twice.
      A     "M 87.4"; // Delivery
      AN    "M 87.5";
      A     "B 15.7"; // Packet on the Edge - Seen by Exit Sens
      S     "M 283.1"; // Packet Seen (Free)
//;
      A     "M 87.5"; // Delivery Done - Exit Sens Clear
      FP    M    283.0; // Edge Memory (Free)
      A     "M 283.1"; // Only if a Packet was Seen
      L     S5T#500MS;
      SE    "Timer 138"; // Count Down Pulse 500mS (> Preset_MIN 300mS)
//;
      A     "Timer 138"; // Counted
      O     "M 87.6"; // Steps Reset
      R     "M 283.1";
//;
      A     "Timer 138";
      =     #BIT1; // Count Down Pulse
      =     #XFER;
//;
      CALL "DE-BOUNCER / COUNTER" (
           Bit_0                    := #BIT0,
           Bit_1                    := #BIT1,
           Transfer_Start           := #XFER,
           Error_Reset              := "M 9.1",
           Space_DX_mS              := 600,
           ReSample_DX              := 85,
           Conveyor_Type            := 2,
           Preset_MIN_mS            := 300,
           LowSpd_Dimension_mS      := 0,
           HighSpd_Dimension_mS     := 0,
           Plc_Scan_mS              := "DB UTILITY".Scan_Cycle_Previous,
           Q_Error                  := #ERROR,
           Word_Count               := "HMI_DB".CONV_23_COUNT,
           IO_DB                    := "DEBOUNCER COUNTER DB".Conveyor_C23_Delivery);

M540: NOP   0;
NETWORK
TITLE =HMI Packet Counters Reset (Same Conditions as FC1206)
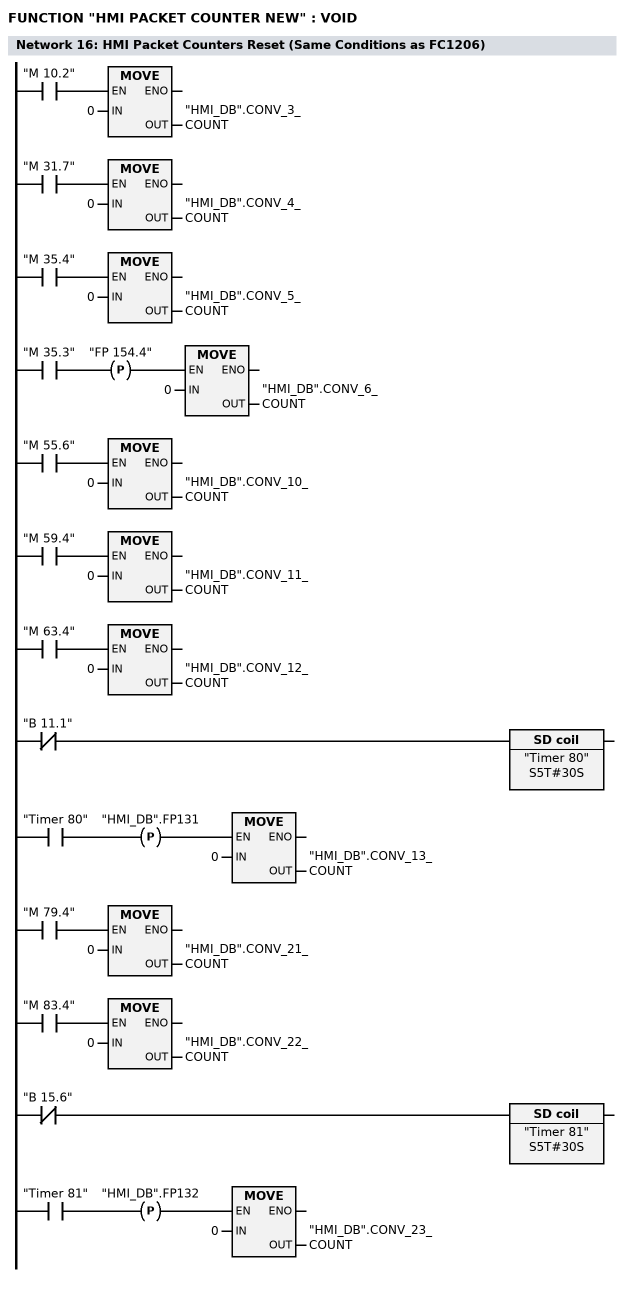

      A     "M 10.2";
      JNB   F102;

      L     0;
      T     "HMI_DB".CONV_3_COUNT; // FC8 Takes Over 0 on Next Call

F102: NOP   0;
      A     "M 31.7";
      JNB   F317;

      L     0;
      T     "HMI_DB".CONV_4_COUNT; // FC8 Takes Over 0 on Next Call

F317: NOP   0;
      A     "M 35.4";
      JNB   F354;

      L     0;
      T     "HMI_DB".CONV_5_COUNT; // FC8 Takes Over 0 on Next Call

F354: NOP   0;
      A     "M 35.3";
      FP    "FP 154.4";
      JNB   F396;

      L     0;
      T     "HMI_DB".CONV_6_COUNT; // FC8 Takes Over 0 on Next Call

F396: NOP   0;
      A     "M 55.6";
      JNB   F556;

      L     0;
      T     "HMI_DB".CONV_10_COUNT; // FC8 Takes Over 0 on Next Call

F556: NOP   0;
      A     "M 59.4";
      JNB   F594;

      L     0;
      T     "HMI_DB".CONV_11_COUNT; // FC8 Takes Over 0 on Next Call

F594: NOP   0;
      A     "M 63.4";
      JNB   F634;

      L     0;
      T     "HMI_DB".CONV_12_COUNT; // FC8 Takes Over 0 on Next Call

F634: NOP   0;
      AN    "B 11.1";
      L     S5T#30S;
      SD    "Timer 80";
//;
      A     "Timer 80";
      FP    "HMI_DB".FP131;
      JNB   F676;

      L     0;
      T     "HMI_DB".CONV_13_COUNT; // FC8 Takes Over 0 on Next Call

F676: NOP   0;
      A     "M 79.4";
      JNB   F794;

      L     0;
      T     "HMI_DB".CONV_21_COUNT; // FC8 Takes Over 0 on Next Call

F794: NOP   0;
      A     "M 83.4";
      JNB   F834;

      L     0;
      T     "HMI_DB".CONV_22_COUNT; // FC8 Takes Over 0 on Next Call

F834: NOP   0;
      AN    "B 15.6";
      L     S5T#30S;
      SD    "Timer 81";
//;
      A     "Timer 81";
      FP    "HMI_DB".FP132;
      JNB   F876;

      L     0;
      T     "HMI_DB".CONV_23_COUNT; // FC8 Takes Over 0 on Next Call

F876: NOP   0;
END_FUNCTION

FUNCTION "PACKET WIDTH MEASURE" : VOID
TITLE =Packet Width Measure - C10 Transfer, B10.5 + B10.6
//MEASUREMENT ONLY (v0.1): writes only "PACKET WIDTH DB" (DB30), changes nothing
//on the machine. While C10 transfers (M55.5), every packet passing B10.5 and
//B10.6 is measured with the C10 encoder (FM350 ch5). At the end of the
//transfer both sensors must agree (same number of packets, = C10 count, and
//average widths within Tolerance_Pct) -> Width_mm (encoder) and Width_ms_31
//(measured, = C11/C12/C13 + C21/C22/C23 loading speed) are VERIFIED.
//v0.9 2026-11-19: direct encoder steps < 0 or > 300 pulses/scan ignored (Ch5
//restarts from 0 when gate 5 reopens).
//v0.8 2026-11-19: also runs the packet BLANKING in shadow (FC1212 / DB31): one
//cleaned count per packet at the C10/C11/C12/C21/C22 exits, NOT used by FC1208
//yet.
VERSION : 0.9


VAR_TEMP
  START : BOOL ;
  STOP : BOOL ;
  OK : BOOL ;
  GAP_P : DINT ;
  C5 : INT ;
  C6 : INT ;
  DIFF : INT ;
  TOLMM : INT ;
  D : DINT ;
  PTR : DWORD ;
  WB : INT ;
  RUNB : BOOL ;
  PLS : BOOL ;
  W : INT ;
  DW : DINT ;
END_VAR
BEGIN
NETWORK
TITLE =C10 Transfer - Start / End
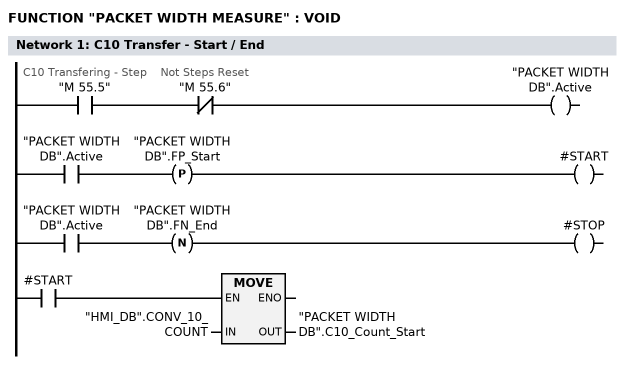

      A     "M 55.5"; // C10 Transfering - Step
      AN    "M 55.6"; // Not Steps Reset
      =     "PACKET WIDTH DB".Active;
//;
      A     "PACKET WIDTH DB".Active;
      FP    "PACKET WIDTH DB".FP_Start;
      =     #START;
//;
      A     "PACKET WIDTH DB".Active;
      FN    "PACKET WIDTH DB".FN_End;
      =     #STOP;
//;
      A     #START;
      JCN   W001;

      L     "HMI_DB".CONV_10_COUNT; // Packets on C10 Before Transfer
      T     "PACKET WIDTH DB".C10_Count_Start;

W001: NOP   0;
NETWORK
TITLE =Gap Minimum mm -> Encoder Pulses

      L     "PACKET WIDTH DB".Gap_Min_mm;
      ITD   ;
      DTR   ;
      L     3.100000e-001;
      /R    ;
      RND   ;
      T     #GAP_P;
NETWORK
TITLE =Encoder Source - Read Job Value or Direct Peripheral Word (Every
//ACT_CNTV5 comes from the CNT2_RD job 101, fired once per 100 mS (M6.0), so it
//can be 100 mS or more old (51 mm @ 30.6 m/min). Direct = PIW of the FM350-2
//direct area (low word of Ch5, every scan). The word wraps at 65536: only the
//difference to the last scan (INT, wrap-safe) is added to Enc_Live (DINT).
      A     "PACKET WIDTH DB".Enc_Direct;
      JCN   E001;

      L     "PACKET WIDTH DB".Enc_PIW_Addr;
      SLD   3; // Byte Address -> Pointer
      T     #PTR;
      L     PIW [#PTR];
      T     #W;
//;
      A     "PACKET WIDTH DB".Enc_Direct_Mem; // First Scan in Direct Mode: Init
      JC    E003;

      L     #W;
      T     "PACKET WIDTH DB".Enc_Word_Last;
      SET   ;
      =     "PACKET WIDTH DB".Enc_Direct_Mem;
      JU    E002;

E003: L     #W; // Pulses Since Last Scan (INT Subtraction = Wrap-Safe)
      L     "PACKET WIDTH DB".Enc_Word_Last;
      -I    ;
      ITD   ;
      T     #DW;
      L     L#0; // Ch5 Restarts from 0 When Gate 5 Reopens: Negative or
      <D    ; // Big Step = Restart, Not Travel -> Ignored
      JC    E004;

      L     #DW;
      L     L#300;
      >D    ;
      JC    E004;

      L     "PACKET WIDTH DB".Enc_Live;
      L     #DW;
      +D    ;
      T     "PACKET WIDTH DB".Enc_Live;

E004: NOP   0;
      L     #W;
      T     "PACKET WIDTH DB".Enc_Word_Last;
      JU    E002;

E001: CLR   ;
      =     "PACKET WIDTH DB".Enc_Direct_Mem;
      L     "FM350 DB".ACT_CNTV5;
      T     "PACKET WIDTH DB".Enc_Live;

E002: NOP   0;
NETWORK
TITLE =B10.5 C10 Full Sens

      CALL "WIDTH SENSOR" (
           Sensor                   := "B 10.5",
           Active                   := "PACKET WIDTH DB".Active,
           Start                    := #START,
           Stop                     := #STOP,
           Enc                      := "PACKET WIDTH DB".Enc_Live,
           Gap_Min_Pulse            := #GAP_P,
           Scan_mS                  := "DB UTILITY".Scan_Cycle_Previous,
           Data                     := "PACKET WIDTH DB".S5);
NETWORK
TITLE =B10.6 C10 Exit Sens

      CALL "WIDTH SENSOR" (
           Sensor                   := "B 10.6",
           Active                   := "PACKET WIDTH DB".Active,
           Start                    := #START,
           Stop                     := #STOP,
           Enc                      := "PACKET WIDTH DB".Enc_Live,
           Gap_Min_Pulse            := #GAP_P,
           Scan_mS                  := "DB UTILITY".Scan_Cycle_Previous,
           Data                     := "PACKET WIDTH DB".S6);
NETWORK
TITLE =Calibration - Same Packet Front at B10.5 then B10.6
//Pitch (packet + gap, ~650 mm) > Sensor_Dist (527 mm): the first front at B10.6
//after a front at B10.5 is the SAME packet. Pulses and mS between the two give
//the real mm/pulse and the real C10 speed - every transfer, no jog needed.
      A     #START;
      JCN   K001;

      L     L#0;
      T     "PACKET WIDTH DB".T_ms;
      T     "PACKET WIDTH DB".Cal_Pulse_Sum;
      T     "PACKET WIDTH DB".Cal_ms_Sum;
      L     0;
      T     "PACKET WIDTH DB".Cal_Count;
      CLR   ;
      =     "PACKET WIDTH DB".Pend;

K001: A     "PACKET WIDTH DB".Active;
      JCN   K090;

      L     "PACKET WIDTH DB".T_ms;
      L     "DB UTILITY".Scan_Cycle_Previous;
      ITD   ;
      +D    ;
      T     "PACKET WIDTH DB".T_ms;
//;
      A     "PACKET WIDTH DB".S6.Front; // B10.6 First (Same Scan Case)
      A     "PACKET WIDTH DB".Pend;
      JCN   K002;

      L     "PACKET WIDTH DB".Enc_Live;
      L     "PACKET WIDTH DB".Pend_Enc;
      -D    ;
      T     #D;
      L     L#0;
      >=D   ;
      JC    K003;

      L     #D;
      NEGD  ;
      T     #D;

K003: L     "PACKET WIDTH DB".Cal_Pulse_Sum;
      L     #D;
      +D    ;
      T     "PACKET WIDTH DB".Cal_Pulse_Sum;
      L     "PACKET WIDTH DB".T_ms;
      L     "PACKET WIDTH DB".Pend_T;
      -D    ;
      L     "PACKET WIDTH DB".Cal_ms_Sum;
      +D    ;
      T     "PACKET WIDTH DB".Cal_ms_Sum;
      L     "PACKET WIDTH DB".Cal_Count;
      L     1;
      +I    ;
      T     "PACKET WIDTH DB".Cal_Count;
      SET   ;
      R     "PACKET WIDTH DB".Pend;

K002: A     "PACKET WIDTH DB".S5.Front;
      JCN   K090;

      L     "PACKET WIDTH DB".Enc_Live;
      T     "PACKET WIDTH DB".Pend_Enc;
      L     "PACKET WIDTH DB".T_ms;
      T     "PACKET WIDTH DB".Pend_T;
      SET   ;
      S     "PACKET WIDTH DB".Pend;

K090: NOP   0;
NETWORK
TITLE =Transfer End - Verify (Both Sensors Agree) and Store

      A     #STOP;
      JCN   W090;

      L     "PACKET WIDTH DB".S5.Count; // Packets Seen = Measured + Partial
      L     "PACKET WIDTH DB".S5.Skipped;
      +I    ;
      T     #C5;
      L     "PACKET WIDTH DB".S6.Count;
      L     "PACKET WIDTH DB".S6.Skipped;
      +I    ;
      T     #C6;
//;
      L     #C5; // No Packet at Both Sensors = Empty Transfer, Not Rejected
      L     0;
      ==I   ;
      A(    ;
      L     #C6;
      L     0;
      ==I   ;
      )     ;
      JCN   W005;

      L     "PACKET WIDTH DB".Empty_Count;
      L     1;
      +I    ;
      T     "PACKET WIDTH DB".Empty_Count;
      JU    W090;

W005: NOP   0;
      L     "PACKET WIDTH DB".S5.Width_Avg_mm;
      L     "PACKET WIDTH DB".S6.Width_Avg_mm;
      -I    ;
      T     #DIFF;
      L     0;
      >=I   ;
      JC    W002;

      L     #DIFF;
      NEGI  ;
      T     #DIFF;

W002: L     "PACKET WIDTH DB".S5.Width_Avg_mm;
      L     "PACKET WIDTH DB".Tolerance_Pct;
      *I    ;
      L     100;
      /I    ;
      T     #TOLMM;
//;
      L     "PACKET WIDTH DB".S5.Count; // Both Measured Something
      L     0;
      >I    ;
      A(    ;
      L     "PACKET WIDTH DB".S6.Count;
      L     0;
      >I    ;
      )     ;
      A(    ;
      L     #C5; // Same Number of Packets
      L     #C6;
      ==I   ;
      )     ;
      A(    ;
      L     #DIFF; // Same Width
      L     #TOLMM;
      <=I   ;
      )     ;
      A(    ;
      L     "PACKET WIDTH DB".C10_Count_Start; // = C10 Count (0 = Unknown)
      L     0;
      ==I   ;
      O     ;
      L     #C5;
      L     "PACKET WIDTH DB".C10_Count_Start;
      ==I   ;
      )     ;
      =     #OK;
      =     "PACKET WIDTH DB".Last_OK;
      JCN   W003;

      L     "PACKET WIDTH DB".S5.Width_Avg_mm;
      L     "PACKET WIDTH DB".S6.Width_Avg_mm;
      +I    ;
      L     2;
      /I    ;
      T     "PACKET WIDTH DB".Width_mm;
//;
      L     "PACKET WIDTH DB".S5.Width_Avg_ms; // MEASURED mS @ C10 Fast
      L     "PACKET WIDTH DB".S6.Width_Avg_ms;
      +I    ;
      L     2;
      /I    ;
      T     "PACKET WIDTH DB".Width_ms_31;
//;
      L     "PACKET WIDTH DB".Width_ms_31; // Check: Speed = mm x 1000 / mS
      L     0;
      >I    ;
      JCN   W004;

      L     "PACKET WIDTH DB".Width_mm;
      ITD   ;
      L     L#1000;
      *D    ;
      L     "PACKET WIDTH DB".Width_ms_31;
      ITD   ;
      /D    ;
      T     "PACKET WIDTH DB".Speed_mm_s;

W004: NOP   0;
      SET   ;
      S     "PACKET WIDTH DB".Valid;
      L     "PACKET WIDTH DB".Good_Count;
      L     1;
      +I    ;
      T     "PACKET WIDTH DB".Good_Count;
      JU    W090;

W003: L     "PACKET WIDTH DB".Bad_Count;
      L     1;
      +I    ;
      T     "PACKET WIDTH DB".Bad_Count;

W090: NOP   0;
NETWORK
TITLE =Transfer End - Calibration Result

      A     #STOP;
      JCN   K190;

      L     "PACKET WIDTH DB".Cal_Count;
      L     0;
      >I    ;
      A(    ;
      L     "PACKET WIDTH DB".Cal_Pulse_Sum;
      L     L#0;
      >D    ;
      )     ;
      A(    ;
      L     "PACKET WIDTH DB".Cal_ms_Sum;
      L     L#0;
      >D    ;
      )     ;
      JCN   K190;

      L     "PACKET WIDTH DB".Sensor_Dist_mm; // mm/pulse = Dist x Count / Pulses
      ITD   ;
      DTR   ;
      L     "PACKET WIDTH DB".Cal_Count;
      ITD   ;
      DTR   ;
      *R    ;
      L     "PACKET WIDTH DB".Cal_Pulse_Sum;
      DTR   ;
      /R    ;
      T     "PACKET WIDTH DB".Cal_mm_Pulse;
//;
      L     "PACKET WIDTH DB".Sensor_Dist_mm; // mm/s = Dist x Count x 1000 / mS
      ITD   ;
      DTR   ;
      L     "PACKET WIDTH DB".Cal_Count;
      ITD   ;
      DTR   ;
      *R    ;
      L     1.000000e+003;
      *R    ;
      L     "PACKET WIDTH DB".Cal_ms_Sum;
      DTR   ;
      /R    ;
      RND   ;
      T     "PACKET WIDTH DB".Cal_Speed_mm_s;
//;
      L     "PACKET WIDTH DB".Width_mm; // Width with the Calibrated Factor
      ITD   ;
      DTR   ;
      L     "PACKET WIDTH DB".Cal_mm_Pulse;
      *R    ;
      L     3.100000e-001;
      /R    ;
      RND   ;
      T     "PACKET WIDTH DB".Width_mm_Cal;

K190: NOP   0;
NETWORK
TITLE =Blanking (Shadow) - Packet Time to Use

      L     "PACKET WIDTH DB".Width_ms_31;
      T     #WB;
      A     "PACKET WIDTH DB".Valid;
      A(    ;
      L     #WB;
      L     300;
      >I    ;
      )     ;
      A(    ;
      L     #WB;
      L     5000;
      <I    ;
      )     ;
      JC    K201;

      L     855; // Default (Measured 2026-11-19)
      T     #WB;

K201: L     #WB;
      T     "BLANKING DB".Width_ms;
NETWORK
TITLE =Blanking (Shadow) - C10 Exit B10.6
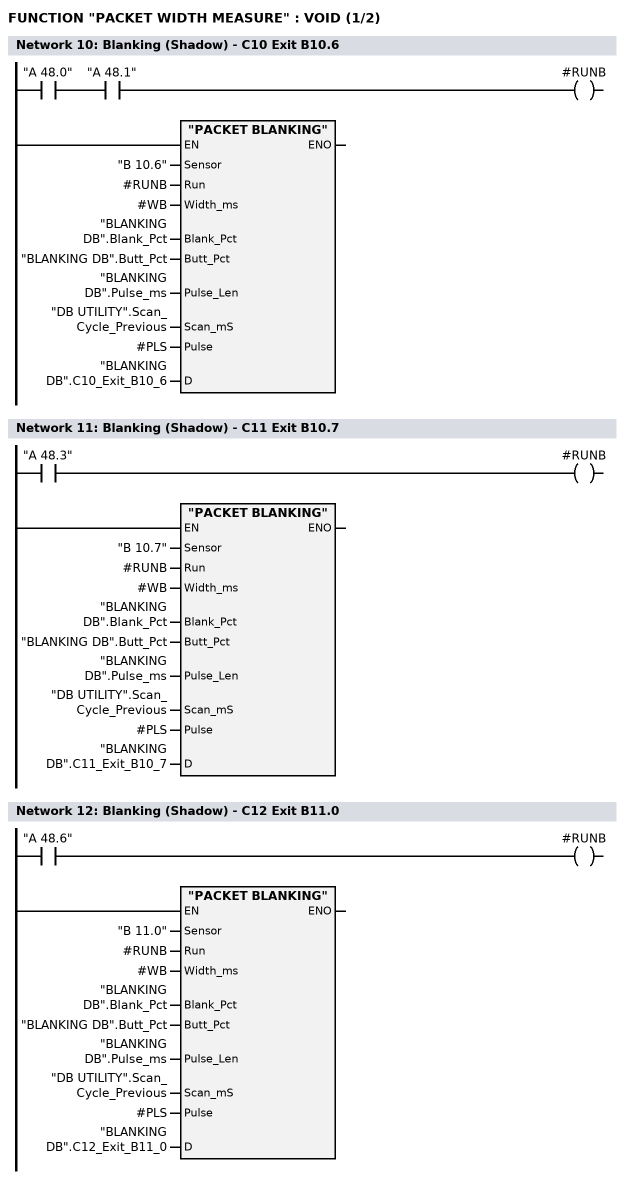

      A     "A 48.0";
      A     "A 48.1";
      =     #RUNB;
      CALL "PACKET BLANKING" (
           Sensor                   := "B 10.6",
           Run                      := #RUNB,
           Width_ms                 := #WB,
           Blank_Pct                := "BLANKING DB".Blank_Pct,
           Butt_Pct                 := "BLANKING DB".Butt_Pct,
           Pulse_Len                := "BLANKING DB".Pulse_ms,
           Scan_mS                  := "DB UTILITY".Scan_Cycle_Previous,
           Pulse                    := #PLS,
           D                        := "BLANKING DB".C10_Exit_B10_6);
NETWORK
TITLE =Blanking (Shadow) - C11 Exit B10.7

      A     "A 48.3";
      =     #RUNB;
      CALL "PACKET BLANKING" (
           Sensor                   := "B 10.7",
           Run                      := #RUNB,
           Width_ms                 := #WB,
           Blank_Pct                := "BLANKING DB".Blank_Pct,
           Butt_Pct                 := "BLANKING DB".Butt_Pct,
           Pulse_Len                := "BLANKING DB".Pulse_ms,
           Scan_mS                  := "DB UTILITY".Scan_Cycle_Previous,
           Pulse                    := #PLS,
           D                        := "BLANKING DB".C11_Exit_B10_7);
NETWORK
TITLE =Blanking (Shadow) - C12 Exit B11.0

      A     "A 48.6";
      =     #RUNB;
      CALL "PACKET BLANKING" (
           Sensor                   := "B 11.0",
           Run                      := #RUNB,
           Width_ms                 := #WB,
           Blank_Pct                := "BLANKING DB".Blank_Pct,
           Butt_Pct                 := "BLANKING DB".Butt_Pct,
           Pulse_Len                := "BLANKING DB".Pulse_ms,
           Scan_mS                  := "DB UTILITY".Scan_Cycle_Previous,
           Pulse                    := #PLS,
           D                        := "BLANKING DB".C12_Exit_B11_0);
NETWORK
TITLE =Blanking (Shadow) - C21 Exit B15.4
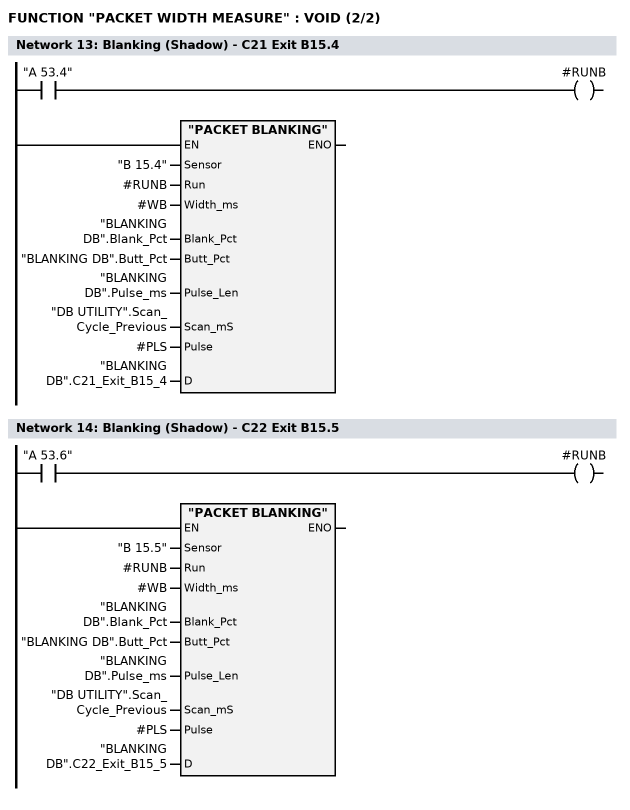

      A     "A 53.4";
      =     #RUNB;
      CALL "PACKET BLANKING" (
           Sensor                   := "B 15.4",
           Run                      := #RUNB,
           Width_ms                 := #WB,
           Blank_Pct                := "BLANKING DB".Blank_Pct,
           Butt_Pct                 := "BLANKING DB".Butt_Pct,
           Pulse_Len                := "BLANKING DB".Pulse_ms,
           Scan_mS                  := "DB UTILITY".Scan_Cycle_Previous,
           Pulse                    := #PLS,
           D                        := "BLANKING DB".C21_Exit_B15_4);
NETWORK
TITLE =Blanking (Shadow) - C22 Exit B15.5

      A     "A 53.6";
      =     #RUNB;
      CALL "PACKET BLANKING" (
           Sensor                   := "B 15.5",
           Run                      := #RUNB,
           Width_ms                 := #WB,
           Blank_Pct                := "BLANKING DB".Blank_Pct,
           Butt_Pct                 := "BLANKING DB".Butt_Pct,
           Pulse_Len                := "BLANKING DB".Pulse_ms,
           Scan_mS                  := "DB UTILITY".Scan_Cycle_Previous,
           Pulse                    := #PLS,
           D                        := "BLANKING DB".C22_Exit_B15_5);
END_FUNCTION

FUNCTION "ALARM MANAGER" : VOID
TITLE =HMI Alarms - NS12 (DB13)
//v1.0 2026-11-23: all LAUER messages (FC199 / FC201) as single alarm bits for
//the NS12 alarm list, ALL at the same time (LAUER showed only the first one).
//Drive faults: one per drive M3.0...M4.7 (LAUER lines for C11 / C21 / C22 / C23
//tested M4.1 = C10 by mistake). Sensor messages: only while the line is empty
//(LAUER cue: M0.3 AND M11.6 AND NOT M9.7), as before.
//Writes only DB13. Changes nothing on the machine.
//v1.1 2026-11-24: + Any_Fault (DBX9.6) / Any_Alarm (DBX9.7) for the NS12 alarm bar.
VERSION : 1.1


VAR_TEMP
  CUE : BOOL ;	//Control ON + Conveyors 1..10 Empty + Clearing Not Done
END_VAR
BEGIN
NETWORK
TITLE =Message Cue (as LAUER MESSAGE1)
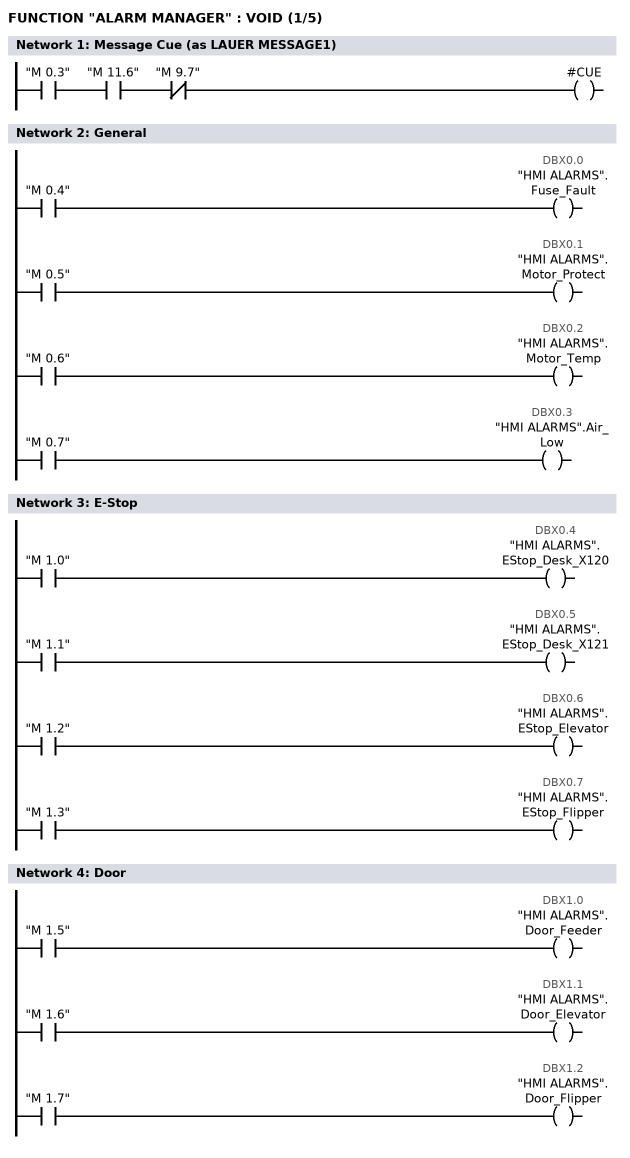

      A     "M 0.3";
      A     "M 11.6";
      AN    "M 9.7";
      =     #CUE;
NETWORK
TITLE =General

      A     "M 0.4";
      =     "HMI ALARMS".Fuse_Fault; // DBX0.0
//;
      A     "M 0.5";
      =     "HMI ALARMS".Motor_Protect; // DBX0.1
//;
      A     "M 0.6";
      =     "HMI ALARMS".Motor_Temp; // DBX0.2
//;
      A     "M 0.7";
      =     "HMI ALARMS".Air_Low; // DBX0.3
NETWORK
TITLE =E-Stop

      A     "M 1.0";
      =     "HMI ALARMS".EStop_Desk_X120; // DBX0.4
//;
      A     "M 1.1";
      =     "HMI ALARMS".EStop_Desk_X121; // DBX0.5
//;
      A     "M 1.2";
      =     "HMI ALARMS".EStop_Elevator; // DBX0.6
//;
      A     "M 1.3";
      =     "HMI ALARMS".EStop_Flipper; // DBX0.7
NETWORK
TITLE =Door

      A     "M 1.5";
      =     "HMI ALARMS".Door_Feeder; // DBX1.0
//;
      A     "M 1.6";
      =     "HMI ALARMS".Door_Elevator; // DBX1.1
//;
      A     "M 1.7";
      =     "HMI ALARMS".Door_Flipper; // DBX1.2
NETWORK
TITLE =Conveyor
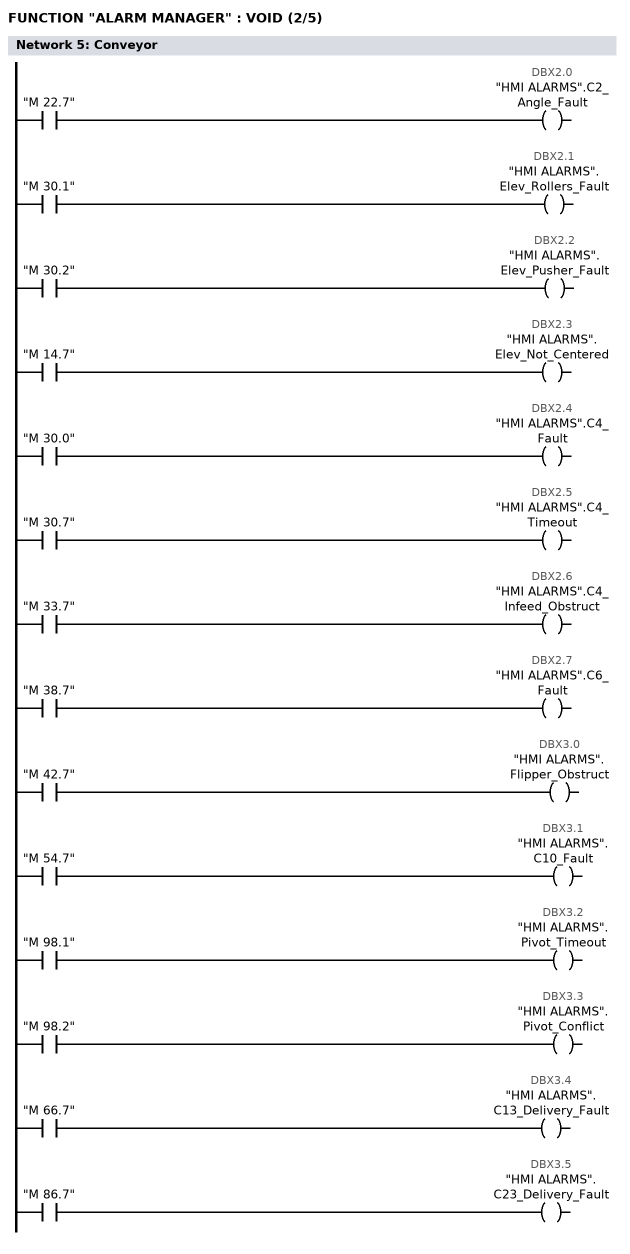

      A     "M 22.7";
      =     "HMI ALARMS".C2_Angle_Fault; // DBX2.0
//;
      A     "M 30.1";
      =     "HMI ALARMS".Elev_Rollers_Fault; // DBX2.1
//;
      A     "M 30.2";
      =     "HMI ALARMS".Elev_Pusher_Fault; // DBX2.2
//;
      A     "M 14.7";
      =     "HMI ALARMS".Elev_Not_Centered; // DBX2.3
//;
      A     "M 30.0";
      =     "HMI ALARMS".C4_Fault; // DBX2.4
//;
      A     "M 30.7";
      =     "HMI ALARMS".C4_Timeout; // DBX2.5
//;
      A     "M 33.7";
      =     "HMI ALARMS".C4_Infeed_Obstruct; // DBX2.6
//;
      A     "M 38.7";
      =     "HMI ALARMS".C6_Fault; // DBX2.7
//;
      A     "M 42.7";
      =     "HMI ALARMS".Flipper_Obstruct; // DBX3.0
//;
      A     "M 54.7";
      =     "HMI ALARMS".C10_Fault; // DBX3.1
//;
      A     "M 98.1";
      =     "HMI ALARMS".Pivot_Timeout; // DBX3.2
//;
      A     "M 98.2";
      =     "HMI ALARMS".Pivot_Conflict; // DBX3.3
//;
      A     "M 66.7";
      =     "HMI ALARMS".C13_Delivery_Fault; // DBX3.4
//;
      A     "M 86.7";
      =     "HMI ALARMS".C23_Delivery_Fault; // DBX3.5
NETWORK
TITLE =Drive
